// --- Siemens Structured Format ---
DATA_BLOCK "model__HS16_IW50_"
{ S7_Optimized_Access := 'TRUE' }
VERSION :
NON_RETAIN
   VAR
      W_i : ARRAY[0..15, 0..39] OF REAL;
      W_f : ARRAY[0..15, 0..39] OF REAL;
      W_g : ARRAY[0..15, 0..39] OF REAL;
      W_o : ARRAY[0..15, 0..39] OF REAL;
      R_i : ARRAY[0..15, 0..15] OF REAL;
      R_f : ARRAY[0..15, 0..15] OF REAL;
      R_g : ARRAY[0..15, 0..15] OF REAL;
      R_o : ARRAY[0..15, 0..15] OF REAL;
      B_i : ARRAY[0..15] OF REAL;
      B_f : ARRAY[0..15] OF REAL;
      B_g : ARRAY[0..15] OF REAL;
      B_o : ARRAY[0..15] OF REAL;
      FC_W : ARRAY[0..39, 0..15] OF REAL;
      FC_B : ARRAY[0..39] OF REAL;
   END_VAR
BEGIN

      W_i[0,0] := -0.02612339;
      W_i[0,1] := 0.12072767;
      W_i[0,2] := -0.02244412;
      W_i[0,3] := -0.02933176;
      W_i[0,4] := 0.13427743;
      W_i[0,5] := -0.01298498;
      W_i[0,6] := -0.08133418;
      W_i[0,7] := 0.19622199;
      W_i[0,8] := 0.14236863;
      W_i[0,9] := -0.06801347;
      W_i[0,10] := 0.16722029;
      W_i[0,11] := -0.33964941;
      W_i[0,12] := -0.82021421;
      W_i[0,13] := 0.06192777;
      W_i[0,14] := 0.39121246;
      W_i[0,15] := -0.96388686;
      W_i[0,16] := 0.14144035;
      W_i[0,17] := -0.25961453;
      W_i[0,18] := 0.00280210;
      W_i[0,19] := 0.36805412;
      W_i[0,20] := 0.11180947;
      W_i[0,21] := 0.28874406;
      W_i[0,22] := 0.24604218;
      W_i[0,23] := 0.06171668;
      W_i[0,24] := 0.88452333;
      W_i[0,25] := 0.96678102;
      W_i[0,26] := 0.04491860;
      W_i[0,27] := -0.21186443;
      W_i[0,28] := 0.08944755;
      W_i[0,29] := -0.10767028;
      W_i[0,30] := 0.60365808;
      W_i[0,31] := -0.13146588;
      W_i[0,32] := 0.12239406;
      W_i[0,33] := -0.09614152;
      W_i[0,34] := 1.05674243;
      W_i[0,35] := -0.04317053;
      W_i[0,36] := 0.15985158;
      W_i[0,37] := -0.00158236;
      W_i[0,38] := 0.64556688;
      W_i[0,39] := 0.15716811;
      W_i[1,0] := 0.02739522;
      W_i[1,1] := 0.10316847;
      W_i[1,2] := 0.01493799;
      W_i[1,3] := 0.01172978;
      W_i[1,4] := 0.17755681;
      W_i[1,5] := 0.02642176;
      W_i[1,6] := 0.08478273;
      W_i[1,7] := 0.04226714;
      W_i[1,8] := 0.00695325;
      W_i[1,9] := 0.03251113;
      W_i[1,10] := 0.02126005;
      W_i[1,11] := -0.01568736;
      W_i[1,12] := -0.09019557;
      W_i[1,13] := -0.08720633;
      W_i[1,14] := 0.02817911;
      W_i[1,15] := -0.01798955;
      W_i[1,16] := -0.04418186;
      W_i[1,17] := 0.01428624;
      W_i[1,18] := -0.27951232;
      W_i[1,19] := 0.05315392;
      W_i[1,20] := -0.10911061;
      W_i[1,21] := 0.05054765;
      W_i[1,22] := 0.18948558;
      W_i[1,23] := -0.08133697;
      W_i[1,24] := -0.40616348;
      W_i[1,25] := -0.53565234;
      W_i[1,26] := -0.10580445;
      W_i[1,27] := -0.17574981;
      W_i[1,28] := -0.05870668;
      W_i[1,29] := 0.05139971;
      W_i[1,30] := 0.03107365;
      W_i[1,31] := -0.09318750;
      W_i[1,32] := -0.25166753;
      W_i[1,33] := -0.11112119;
      W_i[1,34] := 0.15034710;
      W_i[1,35] := -0.26474807;
      W_i[1,36] := -0.05716439;
      W_i[1,37] := -0.00181797;
      W_i[1,38] := 0.06692428;
      W_i[1,39] := -0.00409455;
      W_i[2,0] := -0.04371461;
      W_i[2,1] := 0.03530892;
      W_i[2,2] := -0.03434504;
      W_i[2,3] := -0.05561700;
      W_i[2,4] := 0.00493065;
      W_i[2,5] := 0.03415375;
      W_i[2,6] := -0.02065521;
      W_i[2,7] := -0.04744798;
      W_i[2,8] := 0.11951899;
      W_i[2,9] := 0.11182401;
      W_i[2,10] := 0.04235537;
      W_i[2,11] := -0.08501492;
      W_i[2,12] := 0.08836282;
      W_i[2,13] := -0.03698122;
      W_i[2,14] := 0.11667735;
      W_i[2,15] := -1.35210800;
      W_i[2,16] := 0.04032730;
      W_i[2,17] := 0.39463934;
      W_i[2,18] := 0.23274027;
      W_i[2,19] := -0.09035096;
      W_i[2,20] := 0.02598169;
      W_i[2,21] := -0.02158709;
      W_i[2,22] := 0.08459560;
      W_i[2,23] := -0.01336102;
      W_i[2,24] := 0.39533728;
      W_i[2,25] := 0.21617500;
      W_i[2,26] := 0.04206325;
      W_i[2,27] := 0.03110088;
      W_i[2,28] := 0.00954145;
      W_i[2,29] := -0.08245377;
      W_i[2,30] := -0.01272953;
      W_i[2,31] := -0.00777793;
      W_i[2,32] := -0.03093930;
      W_i[2,33] := -0.14403637;
      W_i[2,34] := -0.36296284;
      W_i[2,35] := 0.02933266;
      W_i[2,36] := 0.00311332;
      W_i[2,37] := 0.06835733;
      W_i[2,38] := 0.13729195;
      W_i[2,39] := -0.09952185;
      W_i[3,0] := 0.00846558;
      W_i[3,1] := -0.12918584;
      W_i[3,2] := -0.00730979;
      W_i[3,3] := 0.01713126;
      W_i[3,4] := -0.02458502;
      W_i[3,5] := -0.01639076;
      W_i[3,6] := -0.17934421;
      W_i[3,7] := -0.01638387;
      W_i[3,8] := -0.03064539;
      W_i[3,9] := 0.08878898;
      W_i[3,10] := -0.07486653;
      W_i[3,11] := -0.08080578;
      W_i[3,12] := 0.06557790;
      W_i[3,13] := 0.01592479;
      W_i[3,14] := -0.03430796;
      W_i[3,15] := 0.01604570;
      W_i[3,16] := 0.01997751;
      W_i[3,17] := -0.03321569;
      W_i[3,18] := 0.04693119;
      W_i[3,19] := 0.00119276;
      W_i[3,20] := -0.06343115;
      W_i[3,21] := 0.07300727;
      W_i[3,22] := 0.17427416;
      W_i[3,23] := -0.07701004;
      W_i[3,24] := -0.04349097;
      W_i[3,25] := 0.08956601;
      W_i[3,26] := -0.03523625;
      W_i[3,27] := -0.00686803;
      W_i[3,28] := -0.01029908;
      W_i[3,29] := 0.05175918;
      W_i[3,30] := 0.10149232;
      W_i[3,31] := -0.11382963;
      W_i[3,32] := 0.07062076;
      W_i[3,33] := -0.01815722;
      W_i[3,34] := 0.04715188;
      W_i[3,35] := -0.06669057;
      W_i[3,36] := 0.01020681;
      W_i[3,37] := 0.25148758;
      W_i[3,38] := -0.01007098;
      W_i[3,39] := -0.00052197;
      W_i[4,0] := 0.06882605;
      W_i[4,1] := 0.29223976;
      W_i[4,2] := 0.13380581;
      W_i[4,3] := -0.35771182;
      W_i[4,4] := 0.25656733;
      W_i[4,5] := -0.20841958;
      W_i[4,6] := 0.07243224;
      W_i[4,7] := 0.38866916;
      W_i[4,8] := 0.53406250;
      W_i[4,9] := -0.23149215;
      W_i[4,10] := -0.19491005;
      W_i[4,11] := -0.48210201;
      W_i[4,12] := 0.13137554;
      W_i[4,13] := 0.50133437;
      W_i[4,14] := -0.01319221;
      W_i[4,15] := -0.16763180;
      W_i[4,16] := -0.02528067;
      W_i[4,17] := 0.20047617;
      W_i[4,18] := 0.07556880;
      W_i[4,19] := 0.12009662;
      W_i[4,20] := -0.23959216;
      W_i[4,21] := -0.05043668;
      W_i[4,22] := 0.03819416;
      W_i[4,23] := 0.32712597;
      W_i[4,24] := -0.06839418;
      W_i[4,25] := -0.00276239;
      W_i[4,26] := -0.26127121;
      W_i[4,27] := -0.20213830;
      W_i[4,28] := 0.07294428;
      W_i[4,29] := 0.04953664;
      W_i[4,30] := -0.04174086;
      W_i[4,31] := -0.06637315;
      W_i[4,32] := 0.09226974;
      W_i[4,33] := 0.13355142;
      W_i[4,34] := 0.09484247;
      W_i[4,35] := -0.09734286;
      W_i[4,36] := 0.03169553;
      W_i[4,37] := -0.08991057;
      W_i[4,38] := -0.13476068;
      W_i[4,39] := 0.29272395;
      W_i[5,0] := -0.05475799;
      W_i[5,1] := -0.06864791;
      W_i[5,2] := -0.02113621;
      W_i[5,3] := 0.02720109;
      W_i[5,4] := 0.10207788;
      W_i[5,5] := -0.00895342;
      W_i[5,6] := -0.02244009;
      W_i[5,7] := 0.16509427;
      W_i[5,8] := 0.01703463;
      W_i[5,9] := -0.21540523;
      W_i[5,10] := -0.00765499;
      W_i[5,11] := 0.01468746;
      W_i[5,12] := 0.22010665;
      W_i[5,13] := -0.09001971;
      W_i[5,14] := -0.02117113;
      W_i[5,15] := 0.07194266;
      W_i[5,16] := -0.18253084;
      W_i[5,17] := 0.04095849;
      W_i[5,18] := -0.08197289;
      W_i[5,19] := -0.27980739;
      W_i[5,20] := 0.11807738;
      W_i[5,21] := 0.25605229;
      W_i[5,22] := -0.18898037;
      W_i[5,23] := 0.06701536;
      W_i[5,24] := -0.38402686;
      W_i[5,25] := 0.03199298;
      W_i[5,26] := 0.28137541;
      W_i[5,27] := -0.03393725;
      W_i[5,28] := -0.00611741;
      W_i[5,29] := -0.21439074;
      W_i[5,30] := -0.24789658;
      W_i[5,31] := 0.01456884;
      W_i[5,32] := 0.09658974;
      W_i[5,33] := 0.07787250;
      W_i[5,34] := -0.00873361;
      W_i[5,35] := 0.02078887;
      W_i[5,36] := -0.00982943;
      W_i[5,37] := -0.22429584;
      W_i[5,38] := 0.25736400;
      W_i[5,39] := -0.30378288;
      W_i[6,0] := -0.15429787;
      W_i[6,1] := -0.00725780;
      W_i[6,2] := -0.01294193;
      W_i[6,3] := -0.08215277;
      W_i[6,4] := -0.13259856;
      W_i[6,5] := -0.16592383;
      W_i[6,6] := -0.00615384;
      W_i[6,7] := 0.02707914;
      W_i[6,8] := 0.03321055;
      W_i[6,9] := 0.20581089;
      W_i[6,10] := -0.02888039;
      W_i[6,11] := 0.13899046;
      W_i[6,12] := -0.50004631;
      W_i[6,13] := -0.18613359;
      W_i[6,14] := 0.02271620;
      W_i[6,15] := -0.05991226;
      W_i[6,16] := 0.02941754;
      W_i[6,17] := -0.05727729;
      W_i[6,18] := -0.05220168;
      W_i[6,19] := 0.12824084;
      W_i[6,20] := -0.11432266;
      W_i[6,21] := -0.06927077;
      W_i[6,22] := -0.16510975;
      W_i[6,23] := 0.16503085;
      W_i[6,24] := -0.06193599;
      W_i[6,25] := 0.08007926;
      W_i[6,26] := 0.16539313;
      W_i[6,27] := -0.09439778;
      W_i[6,28] := -0.11654797;
      W_i[6,29] := -0.07672822;
      W_i[6,30] := -0.09051897;
      W_i[6,31] := -0.05891651;
      W_i[6,32] := -0.06850113;
      W_i[6,33] := -0.01238405;
      W_i[6,34] := 0.05435950;
      W_i[6,35] := -0.07693552;
      W_i[6,36] := 0.00911314;
      W_i[6,37] := -0.01921199;
      W_i[6,38] := 0.05525052;
      W_i[6,39] := -0.07226433;
      W_i[7,0] := -0.19423574;
      W_i[7,1] := -0.24973391;
      W_i[7,2] := -0.05149378;
      W_i[7,3] := -0.25323981;
      W_i[7,4] := 0.39798826;
      W_i[7,5] := 0.24827355;
      W_i[7,6] := 0.43568289;
      W_i[7,7] := -0.13336283;
      W_i[7,8] := 0.12423158;
      W_i[7,9] := -0.07743893;
      W_i[7,10] := -0.15183467;
      W_i[7,11] := 0.06914197;
      W_i[7,12] := -0.02671312;
      W_i[7,13] := -0.21586929;
      W_i[7,14] := 0.00868284;
      W_i[7,15] := 0.02255189;
      W_i[7,16] := -0.02795821;
      W_i[7,17] := 0.00887333;
      W_i[7,18] := -0.12309828;
      W_i[7,19] := -0.00309656;
      W_i[7,20] := 0.38424814;
      W_i[7,21] := 0.30607188;
      W_i[7,22] := -0.15942656;
      W_i[7,23] := 0.01897525;
      W_i[7,24] := -0.09797664;
      W_i[7,25] := -0.02867761;
      W_i[7,26] := 0.15050705;
      W_i[7,27] := 0.00785798;
      W_i[7,28] := -0.19198960;
      W_i[7,29] := 0.21648924;
      W_i[7,30] := 0.16888635;
      W_i[7,31] := -0.00119574;
      W_i[7,32] := -0.24025443;
      W_i[7,33] := 0.30170068;
      W_i[7,34] := 0.23723993;
      W_i[7,35] := -0.13449760;
      W_i[7,36] := -0.15990667;
      W_i[7,37] := -0.00520837;
      W_i[7,38] := 0.08311661;
      W_i[7,39] := -0.02735133;
      W_i[8,0] := -0.06984207;
      W_i[8,1] := 0.18467268;
      W_i[8,2] := 0.00678134;
      W_i[8,3] := 0.04922282;
      W_i[8,4] := 0.11598286;
      W_i[8,5] := 0.08822776;
      W_i[8,6] := -0.10902181;
      W_i[8,7] := -0.16074504;
      W_i[8,8] := -0.11118431;
      W_i[8,9] := 0.10051250;
      W_i[8,10] := 0.07012353;
      W_i[8,11] := 0.07681172;
      W_i[8,12] := -0.22344230;
      W_i[8,13] := -0.12049098;
      W_i[8,14] := 0.01157948;
      W_i[8,15] := 0.01269015;
      W_i[8,16] := 0.01600377;
      W_i[8,17] := 0.02240872;
      W_i[8,18] := -0.02060430;
      W_i[8,19] := -0.06097650;
      W_i[8,20] := 0.07957297;
      W_i[8,21] := 0.08196621;
      W_i[8,22] := -0.02732777;
      W_i[8,23] := -0.06837825;
      W_i[8,24] := -1.24913669;
      W_i[8,25] := -0.21292350;
      W_i[8,26] := 0.05969907;
      W_i[8,27] := -0.15808001;
      W_i[8,28] := -0.06865929;
      W_i[8,29] := -0.05003216;
      W_i[8,30] := 0.13252324;
      W_i[8,31] := -0.10141694;
      W_i[8,32] := 0.15883078;
      W_i[8,33] := 0.01671924;
      W_i[8,34] := 0.01595451;
      W_i[8,35] := 0.04233614;
      W_i[8,36] := 0.10780733;
      W_i[8,37] := 0.00896461;
      W_i[8,38] := 0.13257688;
      W_i[8,39] := 0.05639813;
      W_i[9,0] := 0.04840493;
      W_i[9,1] := 0.00527499;
      W_i[9,2] := -0.03278387;
      W_i[9,3] := 0.08216210;
      W_i[9,4] := -0.01587271;
      W_i[9,5] := -0.00737574;
      W_i[9,6] := -0.01856831;
      W_i[9,7] := 0.19069298;
      W_i[9,8] := -0.00912018;
      W_i[9,9] := -0.24746008;
      W_i[9,10] := -0.06627475;
      W_i[9,11] := 0.07460143;
      W_i[9,12] := -0.04468247;
      W_i[9,13] := -0.03485956;
      W_i[9,14] := -0.02453788;
      W_i[9,15] := 0.00244658;
      W_i[9,16] := -0.00826298;
      W_i[9,17] := 0.00922262;
      W_i[9,18] := 0.03385285;
      W_i[9,19] := 0.04683683;
      W_i[9,20] := -0.03658741;
      W_i[9,21] := -0.05278853;
      W_i[9,22] := -0.06786657;
      W_i[9,23] := -0.03328852;
      W_i[9,24] := -0.67544466;
      W_i[9,25] := -0.45174205;
      W_i[9,26] := 0.01428142;
      W_i[9,27] := 0.00258533;
      W_i[9,28] := -0.00212107;
      W_i[9,29] := 0.26447642;
      W_i[9,30] := -0.04738332;
      W_i[9,31] := 0.02417716;
      W_i[9,32] := -0.13879688;
      W_i[9,33] := 0.05013292;
      W_i[9,34] := -0.61316240;
      W_i[9,35] := -0.11345586;
      W_i[9,36] := -0.00836167;
      W_i[9,37] := 0.06233503;
      W_i[9,38] := -0.01308454;
      W_i[9,39] := 0.00902628;
      W_i[10,0] := 0.05447512;
      W_i[10,1] := 0.00135808;
      W_i[10,2] := 0.00598898;
      W_i[10,3] := -0.00021247;
      W_i[10,4] := 0.00281035;
      W_i[10,5] := -0.01504579;
      W_i[10,6] := 0.12122837;
      W_i[10,7] := -0.06385819;
      W_i[10,8] := -0.04342161;
      W_i[10,9] := 0.08000173;
      W_i[10,10] := 0.01194646;
      W_i[10,11] := 0.11263964;
      W_i[10,12] := 0.04725603;
      W_i[10,13] := -0.02525371;
      W_i[10,14] := 0.01381323;
      W_i[10,15] := 0.00554248;
      W_i[10,16] := -0.01660426;
      W_i[10,17] := 0.00241101;
      W_i[10,18] := 0.01211567;
      W_i[10,19] := 0.01751081;
      W_i[10,20] := -0.00082530;
      W_i[10,21] := 0.03101674;
      W_i[10,22] := -0.26447886;
      W_i[10,23] := 0.02353600;
      W_i[10,24] := -0.22910219;
      W_i[10,25] := -0.38894618;
      W_i[10,26] := -0.03487613;
      W_i[10,27] := -0.11107682;
      W_i[10,28] := -0.06958691;
      W_i[10,29] := 0.15007824;
      W_i[10,30] := 0.10014386;
      W_i[10,31] := 0.07397891;
      W_i[10,32] := -0.12383275;
      W_i[10,33] := 0.08686586;
      W_i[10,34] := -0.85524035;
      W_i[10,35] := 0.14177939;
      W_i[10,36] := -0.02201772;
      W_i[10,37] := 0.01626217;
      W_i[10,38] := 0.16784185;
      W_i[10,39] := 0.00716509;
      W_i[11,0] := -0.08976970;
      W_i[11,1] := -0.00744615;
      W_i[11,2] := -0.05819619;
      W_i[11,3] := -0.07143553;
      W_i[11,4] := -0.03154673;
      W_i[11,5] := 0.03580843;
      W_i[11,6] := -0.03945105;
      W_i[11,7] := -0.12150279;
      W_i[11,8] := 0.00981623;
      W_i[11,9] := 0.05031164;
      W_i[11,10] := -0.02300070;
      W_i[11,11] := -0.08073328;
      W_i[11,12] := 0.01272614;
      W_i[11,13] := -0.07925726;
      W_i[11,14] := 0.00678512;
      W_i[11,15] := 0.04620445;
      W_i[11,16] := -0.00129330;
      W_i[11,17] := 0.00041449;
      W_i[11,18] := 0.03960210;
      W_i[11,19] := -0.01602606;
      W_i[11,20] := 0.02149412;
      W_i[11,21] := -0.02751144;
      W_i[11,22] := -0.15877301;
      W_i[11,23] := 0.01397473;
      W_i[11,24] := -0.66238141;
      W_i[11,25] := -0.94520783;
      W_i[11,26] := -0.10410358;
      W_i[11,27] := -0.01858253;
      W_i[11,28] := -0.07172703;
      W_i[11,29] := 0.25134814;
      W_i[11,30] := -0.14801161;
      W_i[11,31] := -0.01742411;
      W_i[11,32] := 0.07450388;
      W_i[11,33] := -0.03559265;
      W_i[11,34] := -0.21006276;
      W_i[11,35] := 0.20278554;
      W_i[11,36] := -0.01763817;
      W_i[11,37] := -0.27180666;
      W_i[11,38] := 0.05380114;
      W_i[11,39] := 0.00796253;
      W_i[12,0] := 0.25864720;
      W_i[12,1] := -0.12210964;
      W_i[12,2] := -0.14704542;
      W_i[12,3] := -0.03986358;
      W_i[12,4] := 0.08733799;
      W_i[12,5] := -0.37284544;
      W_i[12,6] := 0.10571802;
      W_i[12,7] := -0.11933661;
      W_i[12,8] := -0.06846283;
      W_i[12,9] := 0.08954131;
      W_i[12,10] := -0.22306511;
      W_i[12,11] := 0.46803057;
      W_i[12,12] := 0.21598789;
      W_i[12,13] := -0.09787964;
      W_i[12,14] := 0.15112200;
      W_i[12,15] := 0.20643055;
      W_i[12,16] := -0.07569909;
      W_i[12,17] := -0.00754971;
      W_i[12,18] := -0.09548484;
      W_i[12,19] := 0.01058478;
      W_i[12,20] := 0.47774643;
      W_i[12,21] := -0.12664053;
      W_i[12,22] := 0.20265566;
      W_i[12,23] := 0.19177310;
      W_i[12,24] := 0.31017169;
      W_i[12,25] := 0.23971170;
      W_i[12,26] := -0.31540856;
      W_i[12,27] := 0.03726046;
      W_i[12,28] := -0.08490968;
      W_i[12,29] := 0.18619052;
      W_i[12,30] := 0.18660802;
      W_i[12,31] := -0.07303433;
      W_i[12,32] := 0.10245761;
      W_i[12,33] := -0.12202786;
      W_i[12,34] := -0.00883020;
      W_i[12,35] := -0.27889481;
      W_i[12,36] := 0.19747989;
      W_i[12,37] := -0.33369049;
      W_i[12,38] := 0.28634214;
      W_i[12,39] := 0.08568040;
      W_i[13,0] := -0.12176741;
      W_i[13,1] := 0.13172998;
      W_i[13,2] := -0.01483796;
      W_i[13,3] := -0.02370377;
      W_i[13,4] := 0.14033392;
      W_i[13,5] := -0.02840229;
      W_i[13,6] := -0.06477696;
      W_i[13,7] := -0.09099311;
      W_i[13,8] := -0.02282218;
      W_i[13,9] := 0.24101490;
      W_i[13,10] := 0.02915199;
      W_i[13,11] := -0.20095268;
      W_i[13,12] := -0.41396245;
      W_i[13,13] := -0.09245090;
      W_i[13,14] := 0.02569151;
      W_i[13,15] := -0.04253404;
      W_i[13,16] := -0.03762357;
      W_i[13,17] := 0.03585879;
      W_i[13,18] := 0.01942859;
      W_i[13,19] := 0.13924608;
      W_i[13,20] := 0.02253839;
      W_i[13,21] := 0.04408298;
      W_i[13,22] := 0.11049129;
      W_i[13,23] := 0.09530613;
      W_i[13,24] := 0.22805369;
      W_i[13,25] := -0.03002743;
      W_i[13,26] := 0.14904597;
      W_i[13,27] := 0.04909040;
      W_i[13,28] := -0.01216692;
      W_i[13,29] := -0.08759474;
      W_i[13,30] := 0.09012819;
      W_i[13,31] := -0.05122391;
      W_i[13,32] := -0.07538325;
      W_i[13,33] := 0.01453052;
      W_i[13,34] := -0.06318332;
      W_i[13,35] := -0.08720891;
      W_i[13,36] := 0.07678616;
      W_i[13,37] := 0.13920598;
      W_i[13,38] := -0.06368222;
      W_i[13,39] := 1.11653936;
      W_i[14,0] := -0.07855019;
      W_i[14,1] := 0.03459382;
      W_i[14,2] := -0.02766559;
      W_i[14,3] := 0.04799297;
      W_i[14,4] := 0.02599700;
      W_i[14,5] := 0.06535108;
      W_i[14,6] := 0.00835573;
      W_i[14,7] := -0.06900378;
      W_i[14,8] := -0.02075530;
      W_i[14,9] := 0.05139967;
      W_i[14,10] := 0.01833898;
      W_i[14,11] := -0.09905620;
      W_i[14,12] := 0.04986498;
      W_i[14,13] := 0.08562920;
      W_i[14,14] := 0.04875882;
      W_i[14,15] := 0.21624923;
      W_i[14,16] := -0.09095794;
      W_i[14,17] := -0.00323463;
      W_i[14,18] := 0.52891386;
      W_i[14,19] := -0.31447127;
      W_i[14,20] := 0.04405079;
      W_i[14,21] := -0.04545887;
      W_i[14,22] := -0.18876931;
      W_i[14,23] := -0.04623262;
      W_i[14,24] := -0.37235597;
      W_i[14,25] := -0.34788635;
      W_i[14,26] := -0.16801551;
      W_i[14,27] := 0.07317468;
      W_i[14,28] := 0.02443709;
      W_i[14,29] := 0.24874535;
      W_i[14,30] := -0.39551601;
      W_i[14,31] := -0.07593500;
      W_i[14,32] := -0.28626809;
      W_i[14,33] := -0.31125993;
      W_i[14,34] := -0.64042038;
      W_i[14,35] := 0.03362265;
      W_i[14,36] := 0.02987647;
      W_i[14,37] := -0.11912733;
      W_i[14,38] := 0.20975146;
      W_i[14,39] := 0.74268162;
      W_i[15,0] := 0.05764041;
      W_i[15,1] := 0.01238812;
      W_i[15,2] := -0.00211884;
      W_i[15,3] := -0.15071799;
      W_i[15,4] := -0.05083022;
      W_i[15,5] := 0.03901526;
      W_i[15,6] := -0.02054744;
      W_i[15,7] := 0.00484566;
      W_i[15,8] := 0.03377596;
      W_i[15,9] := 0.06261286;
      W_i[15,10] := 0.02025893;
      W_i[15,11] := 0.09115529;
      W_i[15,12] := 0.02875202;
      W_i[15,13] := 0.02998743;
      W_i[15,14] := -0.00594068;
      W_i[15,15] := -0.01918536;
      W_i[15,16] := -0.01136775;
      W_i[15,17] := 0.00490831;
      W_i[15,18] := -0.07127053;
      W_i[15,19] := -0.02636776;
      W_i[15,20] := 0.06915537;
      W_i[15,21] := 0.25859579;
      W_i[15,22] := -0.39175701;
      W_i[15,23] := 0.03068081;
      W_i[15,24] := -0.66952252;
      W_i[15,25] := -0.82186484;
      W_i[15,26] := 0.00559764;
      W_i[15,27] := -0.04806713;
      W_i[15,28] := -0.05927165;
      W_i[15,29] := -0.02447721;
      W_i[15,30] := -0.35062087;
      W_i[15,31] := -0.01519912;
      W_i[15,32] := -0.12022296;
      W_i[15,33] := 0.17821504;
      W_i[15,34] := -0.81185091;
      W_i[15,35] := -0.22858475;
      W_i[15,36] := -0.06415448;
      W_i[15,37] := -0.17577237;
      W_i[15,38] := 0.00998123;
      W_i[15,39] := 0.04287737;
      W_f[0,0] := 0.04715263;
      W_f[0,1] := 0.10899676;
      W_f[0,2] := -0.06567381;
      W_f[0,3] := 0.08125947;
      W_f[0,4] := -0.12792981;
      W_f[0,5] := 0.02464872;
      W_f[0,6] := -0.00594598;
      W_f[0,7] := 0.00857108;
      W_f[0,8] := -0.02990395;
      W_f[0,9] := -0.03421510;
      W_f[0,10] := 0.10801075;
      W_f[0,11] := -0.16118450;
      W_f[0,12] := 0.06628553;
      W_f[0,13] := -0.00627413;
      W_f[0,14] := -0.09413274;
      W_f[0,15] := -0.02655103;
      W_f[0,16] := 0.04184651;
      W_f[0,17] := -0.13916989;
      W_f[0,18] := -0.11053458;
      W_f[0,19] := -0.15861273;
      W_f[0,20] := 0.03201112;
      W_f[0,21] := 0.19275719;
      W_f[0,22] := 0.27139077;
      W_f[0,23] := -0.01148643;
      W_f[0,24] := 0.96007264;
      W_f[0,25] := 0.87839752;
      W_f[0,26] := -0.03665132;
      W_f[0,27] := -0.01417279;
      W_f[0,28] := -0.03944051;
      W_f[0,29] := -0.21950646;
      W_f[0,30] := 0.28375676;
      W_f[0,31] := 0.06307220;
      W_f[0,32] := 0.33201745;
      W_f[0,33] := 0.12054460;
      W_f[0,34] := 0.68658948;
      W_f[0,35] := 0.23550873;
      W_f[0,36] := -0.01086835;
      W_f[0,37] := -0.08451042;
      W_f[0,38] := -0.00964221;
      W_f[0,39] := -0.03436853;
      W_f[1,0] := 0.08623593;
      W_f[1,1] := -0.73259664;
      W_f[1,2] := 0.08433209;
      W_f[1,3] := -0.03844298;
      W_f[1,4] := -0.11556439;
      W_f[1,5] := 0.20516349;
      W_f[1,6] := -0.10453314;
      W_f[1,7] := -0.04163654;
      W_f[1,8] := -0.04797882;
      W_f[1,9] := -0.06256276;
      W_f[1,10] := -0.09822980;
      W_f[1,11] := 0.12738556;
      W_f[1,12] := 0.23426814;
      W_f[1,13] := 0.09855855;
      W_f[1,14] := 0.03435090;
      W_f[1,15] := 0.11293387;
      W_f[1,16] := -0.19483942;
      W_f[1,17] := -0.03186984;
      W_f[1,18] := 0.66178006;
      W_f[1,19] := 0.02745492;
      W_f[1,20] := 0.35740805;
      W_f[1,21] := -0.25831303;
      W_f[1,22] := -0.12126569;
      W_f[1,23] := 0.22377175;
      W_f[1,24] := -0.83024675;
      W_f[1,25] := -1.25248599;
      W_f[1,26] := 0.28189325;
      W_f[1,27] := -0.13919783;
      W_f[1,28] := -0.02240801;
      W_f[1,29] := -0.18801042;
      W_f[1,30] := -0.04805183;
      W_f[1,31] := 0.24313359;
      W_f[1,32] := 0.26400492;
      W_f[1,33] := 0.17501286;
      W_f[1,34] := 0.51169682;
      W_f[1,35] := 0.40932828;
      W_f[1,36] := -0.35491022;
      W_f[1,37] := -0.03798340;
      W_f[1,38] := -0.08608454;
      W_f[1,39] := 0.02175015;
      W_f[2,0] := -0.00661589;
      W_f[2,1] := -0.13814320;
      W_f[2,2] := 0.02391077;
      W_f[2,3] := 0.15640482;
      W_f[2,4] := 0.00755587;
      W_f[2,5] := -0.04414793;
      W_f[2,6] := -0.05434313;
      W_f[2,7] := 0.06549069;
      W_f[2,8] := -0.15011497;
      W_f[2,9] := -0.08841761;
      W_f[2,10] := 0.00392893;
      W_f[2,11] := 0.61885518;
      W_f[2,12] := 0.55919319;
      W_f[2,13] := 0.02260459;
      W_f[2,14] := -0.20439312;
      W_f[2,15] := 0.25819176;
      W_f[2,16] := 0.00852524;
      W_f[2,17] := 0.36273137;
      W_f[2,18] := -0.45172021;
      W_f[2,19] := 0.06631603;
      W_f[2,20] := 0.09949520;
      W_f[2,21] := 0.06160212;
      W_f[2,22] := -0.03724279;
      W_f[2,23] := -0.01405078;
      W_f[2,24] := -1.01044071;
      W_f[2,25] := -1.24477458;
      W_f[2,26] := 0.06317704;
      W_f[2,27] := -0.12849498;
      W_f[2,28] := -0.01733010;
      W_f[2,29] := 0.30296484;
      W_f[2,30] := -0.06890817;
      W_f[2,31] := 0.12288452;
      W_f[2,32] := 0.03147413;
      W_f[2,33] := 0.24991731;
      W_f[2,34] := 0.14598863;
      W_f[2,35] := -0.05373066;
      W_f[2,36] := -0.08683386;
      W_f[2,37] := 0.17713107;
      W_f[2,38] := -0.31477356;
      W_f[2,39] := 1.00106454;
      W_f[3,0] := -0.00357926;
      W_f[3,1] := -0.02668277;
      W_f[3,2] := -0.02272550;
      W_f[3,3] := 0.04566845;
      W_f[3,4] := -0.05781303;
      W_f[3,5] := -0.05116368;
      W_f[3,6] := 0.33208069;
      W_f[3,7] := 0.05969469;
      W_f[3,8] := 0.04631799;
      W_f[3,9] := -0.07284315;
      W_f[3,10] := 0.02255991;
      W_f[3,11] := 0.05159385;
      W_f[3,12] := -0.20268613;
      W_f[3,13] := 0.01119571;
      W_f[3,14] := -0.05706387;
      W_f[3,15] := -0.07039116;
      W_f[3,16] := 0.01233673;
      W_f[3,17] := -0.11033136;
      W_f[3,18] := 0.03755057;
      W_f[3,19] := -0.15966073;
      W_f[3,20] := -0.00759900;
      W_f[3,21] := 0.02997555;
      W_f[3,22] := -0.00575700;
      W_f[3,23] := 0.09471051;
      W_f[3,24] := -0.76867020;
      W_f[3,25] := -1.10453773;
      W_f[3,26] := 0.08160409;
      W_f[3,27] := 0.07287289;
      W_f[3,28] := -0.23396601;
      W_f[3,29] := -0.01620052;
      W_f[3,30] := -0.14668229;
      W_f[3,31] := 0.29359242;
      W_f[3,32] := 0.28141207;
      W_f[3,33] := 0.10357075;
      W_f[3,34] := 0.15553899;
      W_f[3,35] := -0.08215727;
      W_f[3,36] := 0.59300834;
      W_f[3,37] := 0.06939243;
      W_f[3,38] := 0.05595111;
      W_f[3,39] := -0.01764361;
      W_f[4,0] := -0.04732760;
      W_f[4,1] := 0.14226569;
      W_f[4,2] := -0.19679488;
      W_f[4,3] := 0.03169706;
      W_f[4,4] := 0.03950732;
      W_f[4,5] := 0.12956409;
      W_f[4,6] := -0.13465910;
      W_f[4,7] := -0.11123411;
      W_f[4,8] := 0.01169378;
      W_f[4,9] := -0.00041270;
      W_f[4,10] := 0.06247496;
      W_f[4,11] := -0.19790170;
      W_f[4,12] := -0.13562107;
      W_f[4,13] := 0.40435797;
      W_f[4,14] := 0.03306964;
      W_f[4,15] := -0.17322055;
      W_f[4,16] := -0.05731088;
      W_f[4,17] := -0.06482833;
      W_f[4,18] := 0.09320654;
      W_f[4,19] := 0.24850778;
      W_f[4,20] := -0.18519133;
      W_f[4,21] := 0.12798916;
      W_f[4,22] := 0.14323689;
      W_f[4,23] := -0.01742595;
      W_f[4,24] := 1.63087487;
      W_f[4,25] := 1.71278691;
      W_f[4,26] := -0.17371880;
      W_f[4,27] := 0.04438495;
      W_f[4,28] := 0.10424647;
      W_f[4,29] := 0.17063302;
      W_f[4,30] := 0.42905927;
      W_f[4,31] := 0.27194634;
      W_f[4,32] := -0.01861881;
      W_f[4,33] := -0.02290395;
      W_f[4,34] := 0.25754037;
      W_f[4,35] := 0.41329530;
      W_f[4,36] := -0.09744941;
      W_f[4,37] := 0.27917421;
      W_f[4,38] := 0.01022570;
      W_f[4,39] := 0.21825342;
      W_f[5,0] := -0.12265578;
      W_f[5,1] := 0.11042612;
      W_f[5,2] := 0.03006834;
      W_f[5,3] := -0.26207334;
      W_f[5,4] := 0.00985776;
      W_f[5,5] := -0.02016665;
      W_f[5,6] := -0.03333576;
      W_f[5,7] := 0.15882950;
      W_f[5,8] := -0.27977559;
      W_f[5,9] := 0.25365406;
      W_f[5,10] := -0.03230783;
      W_f[5,11] := -0.21518956;
      W_f[5,12] := -0.23225260;
      W_f[5,13] := 0.04519130;
      W_f[5,14] := 0.00848376;
      W_f[5,15] := -0.03351771;
      W_f[5,16] := 0.09852035;
      W_f[5,17] := -0.09458777;
      W_f[5,18] := 0.02086790;
      W_f[5,19] := 0.13770969;
      W_f[5,20] := -0.04140184;
      W_f[5,21] := 0.09476180;
      W_f[5,22] := 0.41919291;
      W_f[5,23] := -0.14774488;
      W_f[5,24] := 1.13465798;
      W_f[5,25] := 1.46192527;
      W_f[5,26] := -0.06388761;
      W_f[5,27] := 0.03928265;
      W_f[5,28] := 0.03407076;
      W_f[5,29] := -0.51813745;
      W_f[5,30] := 0.24349271;
      W_f[5,31] := 0.01923511;
      W_f[5,32] := 0.05050964;
      W_f[5,33] := -0.03686145;
      W_f[5,34] := 1.16242385;
      W_f[5,35] := 0.04278161;
      W_f[5,36] := -0.03958681;
      W_f[5,37] := 0.17119792;
      W_f[5,38] := 0.04197992;
      W_f[5,39] := 0.22113459;
      W_f[6,0] := -0.05077897;
      W_f[6,1] := 0.12266269;
      W_f[6,2] := -0.15582716;
      W_f[6,3] := -0.07109610;
      W_f[6,4] := 0.01037609;
      W_f[6,5] := 0.03313427;
      W_f[6,6] := 0.05276644;
      W_f[6,7] := -0.06777491;
      W_f[6,8] := 0.02246877;
      W_f[6,9] := -0.12816820;
      W_f[6,10] := 0.01218652;
      W_f[6,11] := -0.06725728;
      W_f[6,12] := 0.11980707;
      W_f[6,13] := -0.03621849;
      W_f[6,14] := 0.23148635;
      W_f[6,15] := -0.05256491;
      W_f[6,16] := 0.28452423;
      W_f[6,17] := -0.04785041;
      W_f[6,18] := 0.00029584;
      W_f[6,19] := -0.33732000;
      W_f[6,20] := -0.01787652;
      W_f[6,21] := 0.04774499;
      W_f[6,22] := 0.32209477;
      W_f[6,23] := -0.11889420;
      W_f[6,24] := 1.09117067;
      W_f[6,25] := 1.12744486;
      W_f[6,26] := -0.07003234;
      W_f[6,27] := 0.01855475;
      W_f[6,28] := -0.00330310;
      W_f[6,29] := -0.26430756;
      W_f[6,30] := 0.21318698;
      W_f[6,31] := 0.04353658;
      W_f[6,32] := 0.27845708;
      W_f[6,33] := 0.02148022;
      W_f[6,34] := 1.27716565;
      W_f[6,35] := -0.13685782;
      W_f[6,36] := -0.05482837;
      W_f[6,37] := 0.09329895;
      W_f[6,38] := 0.06903394;
      W_f[6,39] := -0.18291597;
      W_f[7,0] := -0.06782078;
      W_f[7,1] := -0.41273677;
      W_f[7,2] := -0.23223357;
      W_f[7,3] := -0.13132100;
      W_f[7,4] := -0.00691312;
      W_f[7,5] := 0.61953580;
      W_f[7,6] := 0.74713135;
      W_f[7,7] := -0.13415965;
      W_f[7,8] := -0.70239842;
      W_f[7,9] := -0.12314104;
      W_f[7,10] := -0.26408386;
      W_f[7,11] := -0.04327460;
      W_f[7,12] := 0.06000946;
      W_f[7,13] := -0.08953854;
      W_f[7,14] := -0.01992717;
      W_f[7,15] := -0.03414788;
      W_f[7,16] := -0.10218910;
      W_f[7,17] := -0.02195402;
      W_f[7,18] := -0.15076502;
      W_f[7,19] := -0.14730737;
      W_f[7,20] := 0.04946668;
      W_f[7,21] := 0.36726916;
      W_f[7,22] := -0.01913268;
      W_f[7,23] := -0.20478757;
      W_f[7,24] := -0.07383893;
      W_f[7,25] := 0.03577507;
      W_f[7,26] := -0.36156556;
      W_f[7,27] := 0.10162932;
      W_f[7,28] := 0.08031812;
      W_f[7,29] := 0.03659641;
      W_f[7,30] := -0.06054391;
      W_f[7,31] := 0.01948766;
      W_f[7,32] := 0.22690910;
      W_f[7,33] := 0.09243126;
      W_f[7,34] := 0.36665705;
      W_f[7,35] := -0.18836242;
      W_f[7,36] := 0.08979291;
      W_f[7,37] := -0.03466015;
      W_f[7,38] := 0.17328687;
      W_f[7,39] := 0.01111504;
      W_f[8,0] := -0.10757597;
      W_f[8,1] := 0.18080002;
      W_f[8,2] := -0.18117517;
      W_f[8,3] := 0.05444926;
      W_f[8,4] := -0.03406826;
      W_f[8,5] := 0.03211219;
      W_f[8,6] := 0.04893153;
      W_f[8,7] := 0.00879812;
      W_f[8,8] := 0.05938864;
      W_f[8,9] := -0.05662099;
      W_f[8,10] := 0.05257615;
      W_f[8,11] := -0.27383971;
      W_f[8,12] := -0.06582582;
      W_f[8,13] := 0.00902832;
      W_f[8,14] := 0.01648709;
      W_f[8,15] := -0.32319725;
      W_f[8,16] := 0.18786642;
      W_f[8,17] := -0.08832575;
      W_f[8,18] := 0.05050201;
      W_f[8,19] := -0.14431089;
      W_f[8,20] := -0.07567763;
      W_f[8,21] := -0.01289035;
      W_f[8,22] := -0.01249675;
      W_f[8,23] := -0.01680613;
      W_f[8,24] := 0.68140340;
      W_f[8,25] := 0.89507484;
      W_f[8,26] := -0.06418619;
      W_f[8,27] := 0.07647979;
      W_f[8,28] := 0.03661409;
      W_f[8,29] := -0.14417614;
      W_f[8,30] := -0.04263573;
      W_f[8,31] := 0.03779473;
      W_f[8,32] := 0.05052606;
      W_f[8,33] := 0.06155790;
      W_f[8,34] := 1.02400410;
      W_f[8,35] := -0.17263915;
      W_f[8,36] := 0.00310001;
      W_f[8,37] := -0.04516594;
      W_f[8,38] := -0.01715083;
      W_f[8,39] := 0.20146139;
      W_f[9,0] := 0.15622687;
      W_f[9,1] := 0.10635939;
      W_f[9,2] := -0.72994000;
      W_f[9,3] := -0.14118610;
      W_f[9,4] := -0.14285882;
      W_f[9,5] := 0.16976678;
      W_f[9,6] := 0.04101548;
      W_f[9,7] := 0.27330139;
      W_f[9,8] := -0.28499794;
      W_f[9,9] := -0.18460013;
      W_f[9,10] := 0.00495566;
      W_f[9,11] := -0.10320173;
      W_f[9,12] := -0.06923575;
      W_f[9,13] := 0.01051456;
      W_f[9,14] := -0.04837225;
      W_f[9,15] := -0.07643475;
      W_f[9,16] := 0.09923542;
      W_f[9,17] := -0.00375771;
      W_f[9,18] := -0.02745963;
      W_f[9,19] := 0.00053912;
      W_f[9,20] := -0.08774224;
      W_f[9,21] := 0.14884678;
      W_f[9,22] := 0.02246397;
      W_f[9,23] := 0.02559338;
      W_f[9,24] := -0.25594050;
      W_f[9,25] := -0.34410420;
      W_f[9,26] := 0.00826990;
      W_f[9,27] := -0.00619870;
      W_f[9,28] := 0.02722283;
      W_f[9,29] := -0.04649381;
      W_f[9,30] := 0.32932112;
      W_f[9,31] := -0.01646173;
      W_f[9,32] := 0.16043368;
      W_f[9,33] := 0.15029813;
      W_f[9,34] := -0.59800792;
      W_f[9,35] := 0.31481645;
      W_f[9,36] := -0.03954235;
      W_f[9,37] := -0.10088660;
      W_f[9,38] := 0.07048618;
      W_f[9,39] := -0.02868455;
      W_f[10,0] := -0.08379000;
      W_f[10,1] := -0.16816668;
      W_f[10,2] := 0.01026458;
      W_f[10,3] := -0.05021837;
      W_f[10,4] := -0.08648673;
      W_f[10,5] := 0.05194992;
      W_f[10,6] := -0.04798879;
      W_f[10,7] := -0.00668964;
      W_f[10,8] := -0.01598040;
      W_f[10,9] := -0.19321908;
      W_f[10,10] := -0.00677647;
      W_f[10,11] := -0.11638412;
      W_f[10,12] := -0.05050007;
      W_f[10,13] := -0.05213704;
      W_f[10,14] := -0.18101706;
      W_f[10,15] := 0.02277401;
      W_f[10,16] := 0.02921080;
      W_f[10,17] := 0.00873813;
      W_f[10,18] := 0.06415650;
      W_f[10,19] := -0.08317487;
      W_f[10,20] := -0.02438755;
      W_f[10,21] := -0.16884466;
      W_f[10,22] := 0.27693939;
      W_f[10,23] := 0.00935439;
      W_f[10,24] := 1.43402386;
      W_f[10,25] := 1.74972332;
      W_f[10,26] := 0.01418469;
      W_f[10,27] := 0.14746916;
      W_f[10,28] := 0.17624062;
      W_f[10,29] := 0.38566202;
      W_f[10,30] := 0.24629667;
      W_f[10,31] := -0.06444994;
      W_f[10,32] := 0.02206947;
      W_f[10,33] := 0.01205150;
      W_f[10,34] := 0.64443576;
      W_f[10,35] := 0.17858964;
      W_f[10,36] := 0.02772049;
      W_f[10,37] := 0.09627288;
      W_f[10,38] := -0.00038884;
      W_f[10,39] := 0.09056027;
      W_f[11,0] := 0.04731990;
      W_f[11,1] := 0.07852971;
      W_f[11,2] := 0.04516530;
      W_f[11,3] := 0.08165582;
      W_f[11,4] := -0.00823189;
      W_f[11,5] := 0.03292342;
      W_f[11,6] := 0.08625521;
      W_f[11,7] := 0.03074309;
      W_f[11,8] := -0.06851767;
      W_f[11,9] := -0.02743477;
      W_f[11,10] := 0.00402056;
      W_f[11,11] := 0.01896705;
      W_f[11,12] := 0.02100093;
      W_f[11,13] := 0.04474377;
      W_f[11,14] := -0.03925331;
      W_f[11,15] := -0.01760299;
      W_f[11,16] := -0.05878574;
      W_f[11,17] := -0.00179996;
      W_f[11,18] := 0.01894562;
      W_f[11,19] := 0.01100245;
      W_f[11,20] := -0.08416440;
      W_f[11,21] := 0.08459154;
      W_f[11,22] := -0.07597429;
      W_f[11,23] := -0.02480526;
      W_f[11,24] := -0.30214685;
      W_f[11,25] := -0.06083889;
      W_f[11,26] := 0.05015881;
      W_f[11,27] := -0.01587165;
      W_f[11,28] := -0.00948480;
      W_f[11,29] := 0.16900283;
      W_f[11,30] := 0.01662034;
      W_f[11,31] := -0.04290604;
      W_f[11,32] := -0.15728204;
      W_f[11,33] := 0.18166886;
      W_f[11,34] := 0.06984576;
      W_f[11,35] := 0.02457202;
      W_f[11,36] := 0.02189556;
      W_f[11,37] := -0.02640078;
      W_f[11,38] := 0.00093580;
      W_f[11,39] := 0.04468563;
      W_f[12,0] := 0.13872766;
      W_f[12,1] := 0.36059234;
      W_f[12,2] := 0.18638378;
      W_f[12,3] := 0.38616773;
      W_f[12,4] := 0.18198954;
      W_f[12,5] := -0.01693199;
      W_f[12,6] := 0.51554531;
      W_f[12,7] := 0.66682684;
      W_f[12,8] := -0.49452236;
      W_f[12,9] := 0.56500375;
      W_f[12,10] := -0.31727192;
      W_f[12,11] := -0.16788831;
      W_f[12,12] := -0.09018624;
      W_f[12,13] := -0.02442008;
      W_f[12,14] := -0.06402968;
      W_f[12,15] := -0.11079653;
      W_f[12,16] := 0.23340648;
      W_f[12,17] := -0.03873094;
      W_f[12,18] := -0.35387737;
      W_f[12,19] := -0.13109617;
      W_f[12,20] := -0.02236723;
      W_f[12,21] := -0.25169286;
      W_f[12,22] := 0.04343348;
      W_f[12,23] := -0.14147434;
      W_f[12,24] := 0.09822226;
      W_f[12,25] := 0.07601354;
      W_f[12,26] := 0.13397673;
      W_f[12,27] := -0.16423117;
      W_f[12,28] := 0.20508496;
      W_f[12,29] := -0.19170563;
      W_f[12,30] := -0.21707255;
      W_f[12,31] := 0.19305049;
      W_f[12,32] := -0.00178745;
      W_f[12,33] := -0.02608595;
      W_f[12,34] := 0.07433556;
      W_f[12,35] := -0.07448775;
      W_f[12,36] := -0.12259015;
      W_f[12,37] := 0.05483592;
      W_f[12,38] := -0.02252366;
      W_f[12,39] := -0.13191852;
      W_f[13,0] := 0.05621623;
      W_f[13,1] := 0.02268710;
      W_f[13,2] := -0.02137025;
      W_f[13,3] := -0.03402603;
      W_f[13,4] := -0.00403033;
      W_f[13,5] := 0.05825109;
      W_f[13,6] := 0.02592259;
      W_f[13,7] := 0.01048357;
      W_f[13,8] := -0.00884827;
      W_f[13,9] := -0.07394934;
      W_f[13,10] := 0.01323845;
      W_f[13,11] := 0.11154817;
      W_f[13,12] := 0.19265266;
      W_f[13,13] := 0.09498972;
      W_f[13,14] := -0.01949506;
      W_f[13,15] := 0.01599856;
      W_f[13,16] := -0.04177938;
      W_f[13,17] := -0.01963896;
      W_f[13,18] := 0.06818765;
      W_f[13,19] := -0.10189550;
      W_f[13,20] := -0.00283599;
      W_f[13,21] := -0.02469871;
      W_f[13,22] := -0.04763987;
      W_f[13,23] := -0.05747910;
      W_f[13,24] := 0.62972993;
      W_f[13,25] := 0.50124347;
      W_f[13,26] := -0.15037754;
      W_f[13,27] := -0.02853806;
      W_f[13,28] := 0.03832513;
      W_f[13,29] := 0.01257216;
      W_f[13,30] := 0.03315365;
      W_f[13,31] := 0.00258718;
      W_f[13,32] := 0.23024213;
      W_f[13,33] := 0.01467210;
      W_f[13,34] := 0.52416134;
      W_f[13,35] := -0.07634575;
      W_f[13,36] := 0.00017335;
      W_f[13,37] := -0.06273333;
      W_f[13,38] := 0.01321615;
      W_f[13,39] := 0.01253699;
      W_f[14,0] := 0.05188091;
      W_f[14,1] := 0.09008571;
      W_f[14,2] := -0.06040832;
      W_f[14,3] := -0.15870132;
      W_f[14,4] := 0.01968341;
      W_f[14,5] := -0.02412392;
      W_f[14,6] := 0.00604502;
      W_f[14,7] := 0.00272764;
      W_f[14,8] := -0.02168215;
      W_f[14,9] := -0.08099962;
      W_f[14,10] := 0.01248098;
      W_f[14,11] := 0.04416423;
      W_f[14,12] := 0.01406407;
      W_f[14,13] := -0.03414071;
      W_f[14,14] := 0.00417258;
      W_f[14,15] := -0.15435918;
      W_f[14,16] := 0.11206103;
      W_f[14,17] := -0.05795342;
      W_f[14,18] := 0.20023122;
      W_f[14,19] := 0.25853318;
      W_f[14,20] := -0.04636193;
      W_f[14,21] := 0.05119645;
      W_f[14,22] := 0.01715696;
      W_f[14,23] := 0.00778349;
      W_f[14,24] := -0.25048414;
      W_f[14,25] := -0.59388351;
      W_f[14,26] := 0.12166926;
      W_f[14,27] := -0.01130306;
      W_f[14,28] := 0.02301564;
      W_f[14,29] := 0.03248704;
      W_f[14,30] := 0.04664331;
      W_f[14,31] := 0.05805317;
      W_f[14,32] := 0.02991675;
      W_f[14,33] := 0.12733400;
      W_f[14,34] := -0.05554454;
      W_f[14,35] := -0.04630656;
      W_f[14,36] := -0.04581423;
      W_f[14,37] := 0.15576649;
      W_f[14,38] := -0.03458373;
      W_f[14,39] := 0.07389181;
      W_f[15,0] := -0.02851857;
      W_f[15,1] := 0.12228543;
      W_f[15,2] := 0.04074666;
      W_f[15,3] := -0.16404167;
      W_f[15,4] := 0.03169363;
      W_f[15,5] := -0.04794145;
      W_f[15,6] := -0.02538486;
      W_f[15,7] := 0.09773283;
      W_f[15,8] := -0.00113020;
      W_f[15,9] := 0.00206907;
      W_f[15,10] := 0.00170394;
      W_f[15,11] := -0.18747102;
      W_f[15,12] := 0.13273963;
      W_f[15,13] := 0.00116777;
      W_f[15,14] := -0.01292728;
      W_f[15,15] := -0.05278755;
      W_f[15,16] := 0.02699348;
      W_f[15,17] := 0.06503567;
      W_f[15,18] := -0.08527236;
      W_f[15,19] := -0.36556801;
      W_f[15,20] := 0.04682306;
      W_f[15,21] := 0.18975946;
      W_f[15,22] := 0.58196318;
      W_f[15,23] := 0.01483520;
      W_f[15,24] := 1.57459116;
      W_f[15,25] := 1.53082824;
      W_f[15,26] := 0.08213925;
      W_f[15,27] := 0.17018035;
      W_f[15,28] := 0.16270036;
      W_f[15,29] := -1.25782382;
      W_f[15,30] := 0.78321606;
      W_f[15,31] := -0.03324566;
      W_f[15,32] := 0.06538258;
      W_f[15,33] := 0.22916409;
      W_f[15,34] := 1.10171151;
      W_f[15,35] := 0.06133924;
      W_f[15,36] := -0.06126631;
      W_f[15,37] := 0.05620775;
      W_f[15,38] := 0.02675290;
      W_f[15,39] := 0.08648319;
      W_g[0,0] := -0.03288272;
      W_g[0,1] := 0.06879283;
      W_g[0,2] := -0.02887416;
      W_g[0,3] := 0.02746971;
      W_g[0,4] := 0.04634671;
      W_g[0,5] := -0.01307166;
      W_g[0,6] := 0.04332437;
      W_g[0,7] := 0.02397616;
      W_g[0,8] := 0.02618686;
      W_g[0,9] := 0.02531774;
      W_g[0,10] := -0.00689762;
      W_g[0,11] := -0.03228850;
      W_g[0,12] := -0.04695914;
      W_g[0,13] := -0.00249899;
      W_g[0,14] := -0.06194285;
      W_g[0,15] := -0.01109950;
      W_g[0,16] := 0.00831518;
      W_g[0,17] := -0.11515938;
      W_g[0,18] := 0.00697446;
      W_g[0,19] := -0.06260984;
      W_g[0,20] := -0.06981920;
      W_g[0,21] := -0.10400263;
      W_g[0,22] := 0.00419812;
      W_g[0,23] := 0.02415262;
      W_g[0,24] := -0.13206881;
      W_g[0,25] := 0.14327736;
      W_g[0,26] := 0.07169567;
      W_g[0,27] := -0.13220897;
      W_g[0,28] := 0.07111509;
      W_g[0,29] := 0.00454173;
      W_g[0,30] := -0.00463334;
      W_g[0,31] := 0.00058220;
      W_g[0,32] := 0.00037708;
      W_g[0,33] := -0.00026135;
      W_g[0,34] := 0.22679581;
      W_g[0,35] := 0.00052285;
      W_g[0,36] := 0.00264373;
      W_g[0,37] := -0.02689169;
      W_g[0,38] := -0.00969260;
      W_g[0,39] := -0.03882377;
      W_g[1,0] := -0.05839003;
      W_g[1,1] := 0.42263713;
      W_g[1,2] := -0.04012571;
      W_g[1,3] := 0.01434622;
      W_g[1,4] := -0.05931747;
      W_g[1,5] := -0.09267445;
      W_g[1,6] := 0.09244086;
      W_g[1,7] := 0.00149189;
      W_g[1,8] := 0.01646185;
      W_g[1,9] := 0.00913838;
      W_g[1,10] := 0.01058344;
      W_g[1,11] := -0.03441796;
      W_g[1,12] := -0.02675500;
      W_g[1,13] := -0.01039137;
      W_g[1,14] := -0.02187960;
      W_g[1,15] := -0.03511444;
      W_g[1,16] := 0.06820389;
      W_g[1,17] := 0.00374079;
      W_g[1,18] := 0.09911744;
      W_g[1,19] := -0.02790303;
      W_g[1,20] := -0.21210110;
      W_g[1,21] := 0.14164248;
      W_g[1,22] := -0.04919457;
      W_g[1,23] := -0.10424531;
      W_g[1,24] := -0.25002548;
      W_g[1,25] := -0.41824010;
      W_g[1,26] := -0.05768240;
      W_g[1,27] := 0.16974758;
      W_g[1,28] := 0.08134635;
      W_g[1,29] := 0.01095367;
      W_g[1,30] := -0.10672898;
      W_g[1,31] := -0.03143495;
      W_g[1,32] := -0.05365749;
      W_g[1,33] := 0.00830225;
      W_g[1,34] := 0.00796971;
      W_g[1,35] := -0.11966703;
      W_g[1,36] := 0.10712396;
      W_g[1,37] := 0.04311150;
      W_g[1,38] := 0.02923429;
      W_g[1,39] := 0.00462070;
      W_g[2,0] := -0.01095263;
      W_g[2,1] := 0.07733528;
      W_g[2,2] := -0.00723971;
      W_g[2,3] := 0.00655987;
      W_g[2,4] := 0.05033382;
      W_g[2,5] := -0.05086170;
      W_g[2,6] := -0.00893102;
      W_g[2,7] := 0.00838173;
      W_g[2,8] := 0.01219127;
      W_g[2,9] := -0.00249959;
      W_g[2,10] := 0.01104422;
      W_g[2,11] := 0.08935806;
      W_g[2,12] := 0.05025892;
      W_g[2,13] := 0.01599896;
      W_g[2,14] := -0.14540766;
      W_g[2,15] := 0.03795051;
      W_g[2,16] := 0.00179014;
      W_g[2,17] := 0.12772407;
      W_g[2,18] := -0.09817299;
      W_g[2,19] := 0.13920712;
      W_g[2,20] := 0.00742573;
      W_g[2,21] := 0.00262788;
      W_g[2,22] := 0.01521684;
      W_g[2,23] := -0.00954701;
      W_g[2,24] := 0.62358665;
      W_g[2,25] := 0.38909104;
      W_g[2,26] := 0.02143394;
      W_g[2,27] := 0.01759339;
      W_g[2,28] := 0.06352523;
      W_g[2,29] := -0.04855579;
      W_g[2,30] := 0.02580756;
      W_g[2,31] := 0.00596368;
      W_g[2,32] := 0.01640637;
      W_g[2,33] := 0.02091035;
      W_g[2,34] := 0.49321541;
      W_g[2,35] := 0.03743263;
      W_g[2,36] := -0.01044649;
      W_g[2,37] := -0.00274277;
      W_g[2,38] := 0.00144159;
      W_g[2,39] := -0.59162003;
      W_g[3,0] := -0.02036412;
      W_g[3,1] := -0.14411704;
      W_g[3,2] := -0.02639455;
      W_g[3,3] := 0.02397250;
      W_g[3,4] := -0.16004682;
      W_g[3,5] := -0.00529983;
      W_g[3,6] := 0.13255818;
      W_g[3,7] := 0.02613736;
      W_g[3,8] := 0.01934580;
      W_g[3,9] := 0.02009285;
      W_g[3,10] := -0.06752108;
      W_g[3,11] := -0.04748070;
      W_g[3,12] := -0.05999199;
      W_g[3,13] := 0.00653862;
      W_g[3,14] := -0.03967655;
      W_g[3,15] := -0.03746946;
      W_g[3,16] := 0.02267453;
      W_g[3,17] := -0.07123119;
      W_g[3,18] := 0.03707521;
      W_g[3,19] := -0.06942015;
      W_g[3,20] := -0.10585976;
      W_g[3,21] := 0.07069318;
      W_g[3,22] := 0.04288564;
      W_g[3,23] := 0.09068061;
      W_g[3,24] := 0.25938836;
      W_g[3,25] := -0.00764711;
      W_g[3,26] := -0.00429336;
      W_g[3,27] := 0.10295356;
      W_g[3,28] := -0.12612087;
      W_g[3,29] := 0.00479916;
      W_g[3,30] := 0.15239407;
      W_g[3,31] := 0.05638619;
      W_g[3,32] := 0.05324322;
      W_g[3,33] := 0.03522293;
      W_g[3,34] := 0.02783547;
      W_g[3,35] := -0.00447224;
      W_g[3,36] := 0.34176287;
      W_g[3,37] := 0.15846112;
      W_g[3,38] := 0.02763572;
      W_g[3,39] := -0.00952189;
      W_g[4,0] := 0.05488009;
      W_g[4,1] := -0.00670369;
      W_g[4,2] := 0.04741509;
      W_g[4,3] := 0.00571730;
      W_g[4,4] := -0.06987662;
      W_g[4,5] := 0.01855648;
      W_g[4,6] := 0.09008339;
      W_g[4,7] := 0.00667926;
      W_g[4,8] := 0.00658040;
      W_g[4,9] := 0.00961057;
      W_g[4,10] := -0.04362585;
      W_g[4,11] := -0.03329441;
      W_g[4,12] := -0.01316141;
      W_g[4,13] := 0.14691545;
      W_g[4,14] := 0.00850634;
      W_g[4,15] := -0.05621828;
      W_g[4,16] := -0.05743054;
      W_g[4,17] := 0.13111739;
      W_g[4,18] := 0.00087735;
      W_g[4,19] := -0.02226411;
      W_g[4,20] := -0.11267117;
      W_g[4,21] := -0.02835003;
      W_g[4,22] := -0.02741843;
      W_g[4,23] := 0.13355793;
      W_g[4,24] := -0.16290458;
      W_g[4,25] := -0.17808466;
      W_g[4,26] := 0.02852475;
      W_g[4,27] := -0.02260069;
      W_g[4,28] := 0.03386381;
      W_g[4,29] := 0.04136939;
      W_g[4,30] := -0.02621254;
      W_g[4,31] := -0.02350034;
      W_g[4,32] := -0.02518253;
      W_g[4,33] := -0.02326495;
      W_g[4,34] := -0.32219490;
      W_g[4,35] := -0.05711325;
      W_g[4,36] := 0.05694984;
      W_g[4,37] := 0.00658011;
      W_g[4,38] := -0.06881828;
      W_g[4,39] := -0.02566535;
      W_g[5,0] := -0.12075401;
      W_g[5,1] := 0.02553332;
      W_g[5,2] := -0.12287396;
      W_g[5,3] := 0.12021825;
      W_g[5,4] := -0.07048963;
      W_g[5,5] := -0.14113422;
      W_g[5,6] := 0.05872258;
      W_g[5,7] := 0.12207281;
      W_g[5,8] := 0.11423667;
      W_g[5,9] := 0.12041245;
      W_g[5,10] := 0.01521803;
      W_g[5,11] := -0.01810576;
      W_g[5,12] := -0.00813478;
      W_g[5,13] := -0.08835436;
      W_g[5,14] := 0.09394597;
      W_g[5,15] := -0.04471128;
      W_g[5,16] := -0.06250727;
      W_g[5,17] := 0.06817933;
      W_g[5,18] := -0.01152834;
      W_g[5,19] := -0.00579273;
      W_g[5,20] := -0.08372810;
      W_g[5,21] := -0.06996331;
      W_g[5,22] := 0.01203206;
      W_g[5,23] := 0.00779026;
      W_g[5,24] := 0.08353818;
      W_g[5,25] := -0.25279960;
      W_g[5,26] := 0.05011104;
      W_g[5,27] := -0.10751224;
      W_g[5,28] := -0.07444005;
      W_g[5,29] := -0.02102967;
      W_g[5,30] := 0.00832473;
      W_g[5,31] := 0.01262962;
      W_g[5,32] := -0.01239251;
      W_g[5,33] := 0.00079978;
      W_g[5,34] := 0.07374854;
      W_g[5,35] := -0.04611919;
      W_g[5,36] := -0.01176891;
      W_g[5,37] := 0.02829348;
      W_g[5,38] := 0.00393110;
      W_g[5,39] := 0.07769092;
      W_g[6,0] := -0.05814515;
      W_g[6,1] := -0.04702876;
      W_g[6,2] := -0.06337287;
      W_g[6,3] := 0.03413104;
      W_g[6,4] := 0.06652597;
      W_g[6,5] := -0.05150583;
      W_g[6,6] := -0.01204906;
      W_g[6,7] := 0.03913860;
      W_g[6,8] := 0.03228532;
      W_g[6,9] := 0.03164063;
      W_g[6,10] := 0.01173771;
      W_g[6,11] := -0.01391642;
      W_g[6,12] := -0.03429415;
      W_g[6,13] := -0.04339701;
      W_g[6,14] := 0.06324015;
      W_g[6,15] := -0.00640369;
      W_g[6,16] := 0.18601589;
      W_g[6,17] := -0.00700807;
      W_g[6,18] := 0.00076136;
      W_g[6,19] := -0.05252279;
      W_g[6,20] := 0.04849189;
      W_g[6,21] := 0.02619516;
      W_g[6,22] := -0.00269682;
      W_g[6,23] := -0.02741523;
      W_g[6,24] := 0.05987318;
      W_g[6,25] := 0.04793175;
      W_g[6,26] := -0.02643443;
      W_g[6,27] := 0.04390920;
      W_g[6,28] := 0.03213611;
      W_g[6,29] := 0.01188661;
      W_g[6,30] := -0.01111693;
      W_g[6,31] := -0.00252879;
      W_g[6,32] := -0.00546005;
      W_g[6,33] := -0.00067087;
      W_g[6,34] := 0.17834580;
      W_g[6,35] := 0.00388802;
      W_g[6,36] := -0.02650490;
      W_g[6,37] := 0.01564691;
      W_g[6,38] := -0.30253130;
      W_g[6,39] := -0.15068348;
      W_g[7,0] := -0.10275671;
      W_g[7,1] := -0.24009611;
      W_g[7,2] := -0.11088440;
      W_g[7,3] := -0.01006387;
      W_g[7,4] := -0.03458254;
      W_g[7,5] := 0.23932587;
      W_g[7,6] := 0.40470347;
      W_g[7,7] := -0.00585874;
      W_g[7,8] := -0.01916949;
      W_g[7,9] := -0.00627702;
      W_g[7,10] := -0.27911651;
      W_g[7,11] := 0.01163200;
      W_g[7,12] := 0.01657399;
      W_g[7,13] := -0.10315786;
      W_g[7,14] := 0.03309733;
      W_g[7,15] := 0.00751682;
      W_g[7,16] := -0.02915282;
      W_g[7,17] := 0.03935070;
      W_g[7,18] := -0.12759872;
      W_g[7,19] := 0.04157587;
      W_g[7,20] := -0.30659992;
      W_g[7,21] := 0.09425942;
      W_g[7,22] := -0.00641260;
      W_g[7,23] := -0.09050559;
      W_g[7,24] := 0.01530947;
      W_g[7,25] := -0.15979554;
      W_g[7,26] := -0.00322467;
      W_g[7,27] := 0.04318399;
      W_g[7,28] := 0.14858317;
      W_g[7,29] := 0.04615099;
      W_g[7,30] := 0.00307166;
      W_g[7,31] := 0.04133423;
      W_g[7,32] := 0.00097957;
      W_g[7,33] := 0.02065461;
      W_g[7,34] := 0.04547579;
      W_g[7,35] := -0.00785838;
      W_g[7,36] := -0.20765284;
      W_g[7,37] := 0.00956008;
      W_g[7,38] := 0.00075457;
      W_g[7,39] := 0.02893667;
      W_g[8,0] := -0.08692090;
      W_g[8,1] := 0.08997668;
      W_g[8,2] := -0.09005233;
      W_g[8,3] := -0.01292246;
      W_g[8,4] := 0.10805142;
      W_g[8,5] := 0.14603932;
      W_g[8,6] := -0.02134521;
      W_g[8,7] := -0.01256517;
      W_g[8,8] := -0.01110261;
      W_g[8,9] := -0.01626757;
      W_g[8,10] := 0.05898210;
      W_g[8,11] := -0.11047587;
      W_g[8,12] := -0.09589648;
      W_g[8,13] := -0.02350931;
      W_g[8,14] := 0.02544193;
      W_g[8,15] := -0.13092923;
      W_g[8,16] := 0.10931896;
      W_g[8,17] := 0.12825854;
      W_g[8,18] := 0.12620327;
      W_g[8,19] := -0.12419707;
      W_g[8,20] := 0.03848997;
      W_g[8,21] := -0.06537959;
      W_g[8,22] := 0.00064196;
      W_g[8,23] := -0.03796872;
      W_g[8,24] := -0.04377631;
      W_g[8,25] := -0.30099538;
      W_g[8,26] := 0.02286426;
      W_g[8,27] := -0.06000912;
      W_g[8,28] := 0.03258165;
      W_g[8,29] := -0.02475458;
      W_g[8,30] := -0.00219198;
      W_g[8,31] := -0.00292637;
      W_g[8,32] := 0.00115337;
      W_g[8,33] := 0.00390999;
      W_g[8,34] := -0.04075257;
      W_g[8,35] := -0.02803931;
      W_g[8,36] := 0.02655412;
      W_g[8,37] := 0.02139529;
      W_g[8,38] := 0.04244001;
      W_g[8,39] := 0.03061243;
      W_g[9,0] := -0.22739998;
      W_g[9,1] := -0.12028531;
      W_g[9,2] := -0.22718781;
      W_g[9,3] := -0.18262891;
      W_g[9,4] := -0.01637146;
      W_g[9,5] := -0.23831372;
      W_g[9,6] := 0.00297750;
      W_g[9,7] := -0.17095226;
      W_g[9,8] := -0.18344788;
      W_g[9,9] := -0.18747538;
      W_g[9,10] := -0.31918642;
      W_g[9,11] := -0.01426092;
      W_g[9,12] := -0.00200754;
      W_g[9,13] := 0.00886641;
      W_g[9,14] := -0.01517866;
      W_g[9,15] := -0.00491453;
      W_g[9,16] := 0.03928856;
      W_g[9,17] := 0.05202412;
      W_g[9,18] := -0.04777612;
      W_g[9,19] := 0.00385900;
      W_g[9,20] := 0.04262874;
      W_g[9,21] := -0.05054115;
      W_g[9,22] := -0.04248414;
      W_g[9,23] := -0.00319653;
      W_g[9,24] := -0.31163967;
      W_g[9,25] := -0.09675232;
      W_g[9,26] := -0.01050112;
      W_g[9,27] := -0.05346175;
      W_g[9,28] := -0.06083639;
      W_g[9,29] := 0.12653194;
      W_g[9,30] := -0.05285788;
      W_g[9,31] := -0.01213977;
      W_g[9,32] := -0.04765768;
      W_g[9,33] := -0.05291987;
      W_g[9,34] := -0.29435629;
      W_g[9,35] := -0.06011635;
      W_g[9,36] := -0.05353123;
      W_g[9,37] := 0.00832208;
      W_g[9,38] := 0.00973149;
      W_g[9,39] := -0.01172841;
      W_g[10,0] := 0.03514115;
      W_g[10,1] := 0.11389200;
      W_g[10,2] := 0.03716018;
      W_g[10,3] := -0.01071796;
      W_g[10,4] := -0.30562735;
      W_g[10,5] := 0.01998116;
      W_g[10,6] := 0.14969940;
      W_g[10,7] := -0.02109131;
      W_g[10,8] := -0.01540629;
      W_g[10,9] := -0.00982767;
      W_g[10,10] := -0.09813343;
      W_g[10,11] := -0.09390774;
      W_g[10,12] := -0.09303362;
      W_g[10,13] := -0.00659447;
      W_g[10,14] := -0.08698983;
      W_g[10,15] := -0.09059508;
      W_g[10,16] := -0.01796200;
      W_g[10,17] := -0.02903299;
      W_g[10,18] := 0.13222115;
      W_g[10,19] := -0.13716845;
      W_g[10,20] := -0.15225135;
      W_g[10,21] := 0.03876633;
      W_g[10,22] := 0.04551086;
      W_g[10,23] := 0.02596399;
      W_g[10,24] := 0.15688412;
      W_g[10,25] := 0.16100781;
      W_g[10,26] := 0.01107862;
      W_g[10,27] := -0.07539947;
      W_g[10,28] := -0.25086227;
      W_g[10,29] := -0.12395287;
      W_g[10,30] := 0.05308864;
      W_g[10,31] := 0.06245262;
      W_g[10,32] := 0.03307296;
      W_g[10,33] := 0.04681247;
      W_g[10,34] := 0.23864536;
      W_g[10,35] := 0.01017979;
      W_g[10,36] := -0.34682098;
      W_g[10,37] := 0.01139926;
      W_g[10,38] := -0.06640822;
      W_g[10,39] := -0.07425395;
      W_g[11,0] := -0.20998149;
      W_g[11,1] := 0.05767135;
      W_g[11,2] := -0.23170957;
      W_g[11,3] := 0.02501687;
      W_g[11,4] := 0.02252023;
      W_g[11,5] := 0.03745016;
      W_g[11,6] := 0.00724144;
      W_g[11,7] := 0.03957897;
      W_g[11,8] := 0.02575030;
      W_g[11,9] := 0.03189280;
      W_g[11,10] := 0.05883392;
      W_g[11,11] := 0.02762088;
      W_g[11,12] := 0.01796787;
      W_g[11,13] := 0.28403825;
      W_g[11,14] := 0.06086168;
      W_g[11,15] := 0.02774396;
      W_g[11,16] := 0.03697228;
      W_g[11,17] := -0.07755503;
      W_g[11,18] := -0.01424372;
      W_g[11,19] := 0.01996346;
      W_g[11,20] := 0.13414641;
      W_g[11,21] := 0.12937231;
      W_g[11,22] := -0.01583524;
      W_g[11,23] := 0.26789898;
      W_g[11,24] := 0.32321972;
      W_g[11,25] := 0.31935814;
      W_g[11,26] := -0.05019195;
      W_g[11,27] := 0.23280673;
      W_g[11,28] := 0.09163668;
      W_g[11,29] := -0.01618287;
      W_g[11,30] := -0.00085428;
      W_g[11,31] := -0.01937335;
      W_g[11,32] := 0.01763184;
      W_g[11,33] := -0.00380951;
      W_g[11,34] := 0.07600094;
      W_g[11,35] := 0.09330983;
      W_g[11,36] := -0.07791516;
      W_g[11,37] := 0.01969607;
      W_g[11,38] := 0.04727592;
      W_g[11,39] := 0.04515434;
      W_g[12,0] := -0.05593645;
      W_g[12,1] := -0.04389839;
      W_g[12,2] := -0.05817224;
      W_g[12,3] := 0.04144620;
      W_g[12,4] := -0.02310878;
      W_g[12,5] := 0.04852642;
      W_g[12,6] := -0.08700307;
      W_g[12,7] := 0.03355748;
      W_g[12,8] := 0.03699837;
      W_g[12,9] := 0.03886550;
      W_g[12,10] := 0.10981326;
      W_g[12,11] := -0.09832872;
      W_g[12,12] := -0.09303018;
      W_g[12,13] := -0.04333979;
      W_g[12,14] := -0.11123282;
      W_g[12,15] := -0.09018178;
      W_g[12,16] := -0.00510190;
      W_g[12,17] := -0.01573442;
      W_g[12,18] := -0.70857680;
      W_g[12,19] := -0.04782427;
      W_g[12,20] := 0.08851119;
      W_g[12,21] := 0.02074307;
      W_g[12,22] := -0.01258304;
      W_g[12,23] := -0.00788189;
      W_g[12,24] := -0.11268676;
      W_g[12,25] := -0.11553165;
      W_g[12,26] := -0.01619464;
      W_g[12,27] := 0.04248659;
      W_g[12,28] := -0.07553757;
      W_g[12,29] := 0.02218230;
      W_g[12,30] := -0.02093006;
      W_g[12,31] := -0.01882189;
      W_g[12,32] := -0.01577668;
      W_g[12,33] := -0.00407436;
      W_g[12,34] := -0.14571649;
      W_g[12,35] := -0.03193094;
      W_g[12,36] := 0.03408330;
      W_g[12,37] := -0.00389380;
      W_g[12,38] := 0.02884003;
      W_g[12,39] := -0.03945985;
      W_g[13,0] := 0.04027861;
      W_g[13,1] := -0.07311103;
      W_g[13,2] := 0.04157875;
      W_g[13,3] := 0.01889602;
      W_g[13,4] := -0.11995003;
      W_g[13,5] := -0.01993360;
      W_g[13,6] := 0.03187145;
      W_g[13,7] := 0.01748616;
      W_g[13,8] := 0.01463885;
      W_g[13,9] := 0.02840340;
      W_g[13,10] := -0.02596055;
      W_g[13,11] := 0.02591357;
      W_g[13,12] := 0.02623175;
      W_g[13,13] := -0.00677697;
      W_g[13,14] := -0.00711890;
      W_g[13,15] := 0.05769501;
      W_g[13,16] := 0.30919826;
      W_g[13,17] := 0.02394222;
      W_g[13,18] := -0.03814467;
      W_g[13,19] := 0.01873361;
      W_g[13,20] := -0.05235977;
      W_g[13,21] := -0.04417822;
      W_g[13,22] := -0.01057172;
      W_g[13,23] := 0.04463968;
      W_g[13,24] := 0.05050629;
      W_g[13,25] := -0.15972561;
      W_g[13,26] := 0.02774286;
      W_g[13,27] := -0.08080220;
      W_g[13,28] := -0.09933943;
      W_g[13,29] := 0.03062030;
      W_g[13,30] := -0.00385746;
      W_g[13,31] := 0.01280402;
      W_g[13,32] := -0.00358380;
      W_g[13,33] := -0.00492619;
      W_g[13,34] := 0.04224548;
      W_g[13,35] := -0.00044207;
      W_g[13,36] := -0.04630874;
      W_g[13,37] := -0.03753048;
      W_g[13,38] := 0.09008476;
      W_g[13,39] := 0.02002463;
      W_g[14,0] := 0.06269035;
      W_g[14,1] := 0.16204342;
      W_g[14,2] := 0.07219669;
      W_g[14,3] := -0.04503014;
      W_g[14,4] := -0.00555789;
      W_g[14,5] := 0.01761685;
      W_g[14,6] := -0.03159415;
      W_g[14,7] := -0.05064076;
      W_g[14,8] := -0.04640801;
      W_g[14,9] := -0.06009993;
      W_g[14,10] := 0.00660122;
      W_g[14,11] := -0.03258261;
      W_g[14,12] := -0.03601762;
      W_g[14,13] := 0.03453247;
      W_g[14,14] := 0.12738688;
      W_g[14,15] := -0.01328611;
      W_g[14,16] := 0.01626320;
      W_g[14,17] := -0.04504346;
      W_g[14,18] := -0.15708502;
      W_g[14,19] := 0.00090277;
      W_g[14,20] := -0.04051626;
      W_g[14,21] := -0.04047279;
      W_g[14,22] := 0.00840584;
      W_g[14,23] := -0.01122396;
      W_g[14,24] := 0.06744422;
      W_g[14,25] := 0.49537152;
      W_g[14,26] := 0.07856539;
      W_g[14,27] := -0.03960157;
      W_g[14,28] := 0.03958257;
      W_g[14,29] := -0.04088740;
      W_g[14,30] := 0.02040378;
      W_g[14,31] := 0.01003806;
      W_g[14,32] := 0.02256208;
      W_g[14,33] := 0.02816826;
      W_g[14,34] := 0.15040024;
      W_g[14,35] := 0.01636149;
      W_g[14,36] := 0.04578492;
      W_g[14,37] := -0.03131405;
      W_g[14,38] := -0.05991198;
      W_g[14,39] := 0.01529666;
      W_g[15,0] := 0.11327556;
      W_g[15,1] := -0.17608264;
      W_g[15,2] := 0.09651362;
      W_g[15,3] := 0.02762307;
      W_g[15,4] := 0.26826185;
      W_g[15,5] := -0.27072880;
      W_g[15,6] := 0.04821723;
      W_g[15,7] := 0.03941977;
      W_g[15,8] := 0.02793526;
      W_g[15,9] := 0.03359088;
      W_g[15,10] := -0.12275329;
      W_g[15,11] := -0.16014972;
      W_g[15,12] := -0.16786559;
      W_g[15,13] := 0.09324758;
      W_g[15,14] := -0.00898216;
      W_g[15,15] := -0.16123867;
      W_g[15,16] := 0.02021289;
      W_g[15,17] := -0.01648896;
      W_g[15,18] := -0.00597759;
      W_g[15,19] := -0.16053081;
      W_g[15,20] := 0.04093139;
      W_g[15,21] := 0.06445049;
      W_g[15,22] := 0.04804592;
      W_g[15,23] := 0.06335551;
      W_g[15,24] := 0.06702932;
      W_g[15,25] := 0.00881007;
      W_g[15,26] := 0.00152106;
      W_g[15,27] := 0.07652006;
      W_g[15,28] := 0.30222309;
      W_g[15,29] := -0.08014103;
      W_g[15,30] := 0.06666484;
      W_g[15,31] := 0.00829429;
      W_g[15,32] := 0.10078011;
      W_g[15,33] := 0.06581395;
      W_g[15,34] := 0.08893893;
      W_g[15,35] := 0.15266605;
      W_g[15,36] := -0.17053175;
      W_g[15,37] := -0.07062726;
      W_g[15,38] := 0.07771596;
      W_g[15,39] := 0.04211254;
      W_o[0,0] := 0.12198126;
      W_o[0,1] := 0.14187956;
      W_o[0,2] := -0.01325197;
      W_o[0,3] := -0.07755501;
      W_o[0,4] := -0.21710020;
      W_o[0,5] := 0.13306709;
      W_o[0,6] := -0.10178271;
      W_o[0,7] := -0.14437862;
      W_o[0,8] := 0.02041168;
      W_o[0,9] := 0.04337119;
      W_o[0,10] := 0.22460431;
      W_o[0,11] := -0.27840534;
      W_o[0,12] := 0.35424832;
      W_o[0,13] := 0.20462060;
      W_o[0,14] := -0.34063420;
      W_o[0,15] := 0.18119343;
      W_o[0,16] := -0.08057553;
      W_o[0,17] := -0.48889911;
      W_o[0,18] := 0.81621987;
      W_o[0,19] := 0.08914678;
      W_o[0,20] := 0.22458921;
      W_o[0,21] := 0.74807531;
      W_o[0,22] := 0.98743701;
      W_o[0,23] := -0.22151884;
      W_o[0,24] := 1.91302598;
      W_o[0,25] := 2.06443334;
      W_o[0,26] := -0.67687452;
      W_o[0,27] := -0.00083833;
      W_o[0,28] := -0.11211787;
      W_o[0,29] := -0.28486133;
      W_o[0,30] := 0.70833492;
      W_o[0,31] := 0.04462677;
      W_o[0,32] := 0.38353100;
      W_o[0,33] := 0.09996076;
      W_o[0,34] := 1.72650719;
      W_o[0,35] := 0.41856179;
      W_o[0,36] := 0.03231431;
      W_o[0,37] := 0.25164288;
      W_o[0,38] := 0.06612357;
      W_o[0,39] := -0.00002071;
      W_o[1,0] := -0.03910590;
      W_o[1,1] := 0.27588379;
      W_o[1,2] := 0.10975786;
      W_o[1,3] := -0.09756759;
      W_o[1,4] := -0.59621233;
      W_o[1,5] := -0.42031246;
      W_o[1,6] := -0.09698014;
      W_o[1,7] := 0.15754665;
      W_o[1,8] := -0.00284551;
      W_o[1,9] := 0.02527599;
      W_o[1,10] := -0.01773636;
      W_o[1,11] := -0.30956084;
      W_o[1,12] := 0.23456147;
      W_o[1,13] := 0.24187891;
      W_o[1,14] := 0.16774826;
      W_o[1,15] := 0.13618931;
      W_o[1,16] := -0.05666412;
      W_o[1,17] := -0.01989032;
      W_o[1,18] := -0.31193376;
      W_o[1,19] := -0.24264094;
      W_o[1,20] := -0.49747720;
      W_o[1,21] := 0.33921909;
      W_o[1,22] := -0.08854222;
      W_o[1,23] := 0.46807775;
      W_o[1,24] := -0.29946747;
      W_o[1,25] := -0.03667294;
      W_o[1,26] := 0.20074379;
      W_o[1,27] := 0.39029807;
      W_o[1,28] := -0.37250715;
      W_o[1,29] := -0.00592554;
      W_o[1,30] := -0.22806711;
      W_o[1,31] := -0.08731094;
      W_o[1,32] := -0.04087760;
      W_o[1,33] := 0.00680849;
      W_o[1,34] := -0.19797693;
      W_o[1,35] := -0.33509916;
      W_o[1,36] := 0.24450488;
      W_o[1,37] := -0.10827561;
      W_o[1,38] := 0.90532941;
      W_o[1,39] := 0.24546179;
      W_o[2,0] := -0.00616825;
      W_o[2,1] := 0.13651501;
      W_o[2,2] := -0.09869462;
      W_o[2,3] := -0.07334173;
      W_o[2,4] := -0.02211194;
      W_o[2,5] := 0.05619258;
      W_o[2,6] := 0.10801718;
      W_o[2,7] := 0.14577843;
      W_o[2,8] := 0.09542450;
      W_o[2,9] := 0.04769905;
      W_o[2,10] := 0.04124768;
      W_o[2,11] := -0.33887896;
      W_o[2,12] := 0.43093050;
      W_o[2,13] := 0.04022788;
      W_o[2,14] := 0.01084119;
      W_o[2,15] := 0.23125160;
      W_o[2,16] := 0.00388798;
      W_o[2,17] := -0.03658837;
      W_o[2,18] := -0.47197291;
      W_o[2,19] := 0.30483419;
      W_o[2,20] := -0.05675438;
      W_o[2,21] := -0.20610483;
      W_o[2,22] := -0.15346101;
      W_o[2,23] := -0.01675959;
      W_o[2,24] := -0.10398360;
      W_o[2,25] := 0.05681018;
      W_o[2,26] := -0.06196046;
      W_o[2,27] := 0.19941610;
      W_o[2,28] := 0.04805862;
      W_o[2,29] := 0.23355408;
      W_o[2,30] := -0.05858275;
      W_o[2,31] := -0.03168040;
      W_o[2,32] := -0.18688639;
      W_o[2,33] := 0.00733624;
      W_o[2,34] := 0.03196214;
      W_o[2,35] := -0.02429556;
      W_o[2,36] := -0.04773033;
      W_o[2,37] := -0.08787826;
      W_o[2,38] := 0.01416256;
      W_o[2,39] := 0.77567047;
      W_o[3,0] := 0.21000762;
      W_o[3,1] := 0.56502008;
      W_o[3,2] := 0.01591207;
      W_o[3,3] := -0.11321840;
      W_o[3,4] := 0.23269446;
      W_o[3,5] := 0.09338996;
      W_o[3,6] := 0.12135104;
      W_o[3,7] := 0.30009910;
      W_o[3,8] := 0.28139746;
      W_o[3,9] := -0.11283773;
      W_o[3,10] := -0.12950897;
      W_o[3,11] := -0.16686824;
      W_o[3,12] := 0.02030786;
      W_o[3,13] := 0.21336913;
      W_o[3,14] := -0.06828818;
      W_o[3,15] := -0.10707476;
      W_o[3,16] := 0.01645426;
      W_o[3,17] := -0.08346992;
      W_o[3,18] := 0.58030689;
      W_o[3,19] := 0.02444929;
      W_o[3,20] := -0.22163415;
      W_o[3,21] := 0.61291105;
      W_o[3,22] := -0.28959793;
      W_o[3,23] := -0.06618109;
      W_o[3,24] := 0.31345260;
      W_o[3,25] := 0.13633017;
      W_o[3,26] := -0.08859906;
      W_o[3,27] := -0.25854555;
      W_o[3,28] := -0.18073046;
      W_o[3,29] := -0.06065677;
      W_o[3,30] := -0.42247161;
      W_o[3,31] := 0.19295032;
      W_o[3,32] := -0.42941913;
      W_o[3,33] := 0.22519505;
      W_o[3,34] := -0.16697113;
      W_o[3,35] := -0.12213719;
      W_o[3,36] := 0.07402483;
      W_o[3,37] := -0.18623771;
      W_o[3,38] := -0.06633836;
      W_o[3,39] := -0.00843535;
      W_o[4,0] := -0.08241624;
      W_o[4,1] := -0.15822247;
      W_o[4,2] := -0.10238844;
      W_o[4,3] := -0.03743736;
      W_o[4,4] := 0.04915955;
      W_o[4,5] := 0.13049453;
      W_o[4,6] := 0.17377743;
      W_o[4,7] := -0.06675444;
      W_o[4,8] := -0.03882149;
      W_o[4,9] := 0.06404497;
      W_o[4,10] := 0.00192631;
      W_o[4,11] := -0.45325428;
      W_o[4,12] := 0.25542077;
      W_o[4,13] := -0.36887005;
      W_o[4,14] := -0.18856272;
      W_o[4,15] := -0.13098666;
      W_o[4,16] := -0.22178020;
      W_o[4,17] := -0.29496050;
      W_o[4,18] := -0.00731075;
      W_o[4,19] := -0.09241781;
      W_o[4,20] := -0.26850891;
      W_o[4,21] := -0.20041393;
      W_o[4,22] := -0.53797185;
      W_o[4,23] := 0.50577527;
      W_o[4,24] := 0.98513478;
      W_o[4,25] := 1.10475135;
      W_o[4,26] := 0.09366516;
      W_o[4,27] := 0.19566087;
      W_o[4,28] := -0.13328505;
      W_o[4,29] := 0.94272023;
      W_o[4,30] := -0.46258932;
      W_o[4,31] := -0.09195930;
      W_o[4,32] := -0.36374816;
      W_o[4,33] := -0.29488632;
      W_o[4,34] := 0.08194333;
      W_o[4,35] := -0.11618637;
      W_o[4,36] := -0.10650394;
      W_o[4,37] := -0.00409420;
      W_o[4,38] := 0.08796127;
      W_o[4,39] := 0.13779099;
      W_o[5,0] := 0.00298015;
      W_o[5,1] := 0.14726847;
      W_o[5,2] := -0.24877922;
      W_o[5,3] := 0.03818390;
      W_o[5,4] := 0.25190380;
      W_o[5,5] := 0.09698023;
      W_o[5,6] := 0.03788623;
      W_o[5,7] := -0.32500836;
      W_o[5,8] := -0.47933936;
      W_o[5,9] := -0.17586684;
      W_o[5,10] := 0.30961692;
      W_o[5,11] := -0.56706995;
      W_o[5,12] := -0.13458350;
      W_o[5,13] := 0.30265138;
      W_o[5,14] := 0.28882200;
      W_o[5,15] := -0.02685931;
      W_o[5,16] := 0.24619135;
      W_o[5,17] := 0.35931662;
      W_o[5,18] := 0.34230548;
      W_o[5,19] := 0.21314520;
      W_o[5,20] := 0.00126743;
      W_o[5,21] := 0.08332776;
      W_o[5,22] := 0.14433613;
      W_o[5,23] := -0.15501527;
      W_o[5,24] := 1.35550761;
      W_o[5,25] := 1.45758998;
      W_o[5,26] := -0.42872009;
      W_o[5,27] := 0.11975341;
      W_o[5,28] := 0.12516311;
      W_o[5,29] := -0.25945181;
      W_o[5,30] := 0.03064806;
      W_o[5,31] := -0.06416538;
      W_o[5,32] := 0.31372464;
      W_o[5,33] := 0.25143003;
      W_o[5,34] := 1.32014525;
      W_o[5,35] := 0.40504000;
      W_o[5,36] := 0.00424331;
      W_o[5,37] := 0.38437104;
      W_o[5,38] := 2.31802607;
      W_o[5,39] := 0.42288464;
      W_o[6,0] := 0.16465783;
      W_o[6,1] := -0.00748923;
      W_o[6,2] := -0.15153547;
      W_o[6,3] := -0.01711627;
      W_o[6,4] := -0.16756265;
      W_o[6,5] := 0.34808365;
      W_o[6,6] := 0.00590673;
      W_o[6,7] := -0.27918947;
      W_o[6,8] := 0.17359419;
      W_o[6,9] := 0.49527067;
      W_o[6,10] := -0.00244592;
      W_o[6,11] := -0.14789435;
      W_o[6,12] := 0.29600164;
      W_o[6,13] := -0.48868799;
      W_o[6,14] := -0.21440262;
      W_o[6,15] := -0.28105071;
      W_o[6,16] := 0.27140900;
      W_o[6,17] := -0.17575939;
      W_o[6,18] := 0.43315357;
      W_o[6,19] := 0.25442523;
      W_o[6,20] := 0.02021864;
      W_o[6,21] := 0.36727905;
      W_o[6,22] := 0.55856705;
      W_o[6,23] := 0.36519867;
      W_o[6,24] := 1.27994967;
      W_o[6,25] := 1.31188405;
      W_o[6,26] := 0.44206235;
      W_o[6,27] := 0.09447443;
      W_o[6,28] := 0.11994729;
      W_o[6,29] := -0.26271847;
      W_o[6,30] := 0.48323816;
      W_o[6,31] := -0.07709061;
      W_o[6,32] := 0.14690454;
      W_o[6,33] := 0.00670793;
      W_o[6,34] := 1.35142434;
      W_o[6,35] := 0.04027350;
      W_o[6,36] := 0.06238577;
      W_o[6,37] := 0.32636163;
      W_o[6,38] := -0.25480887;
      W_o[6,39] := 1.13409173;
      W_o[7,0] := 0.07718845;
      W_o[7,1] := 0.20402764;
      W_o[7,2] := 0.06463404;
      W_o[7,3] := 0.02887609;
      W_o[7,4] := -0.05794537;
      W_o[7,5] := 0.19518182;
      W_o[7,6] := 1.15763307;
      W_o[7,7] := 0.05626965;
      W_o[7,8] := 0.02816673;
      W_o[7,9] := 0.21392144;
      W_o[7,10] := -0.00420654;
      W_o[7,11] := -0.07277058;
      W_o[7,12] := 0.01088039;
      W_o[7,13] := 0.02142877;
      W_o[7,14] := -0.03849939;
      W_o[7,15] := -0.00698312;
      W_o[7,16] := 0.03512425;
      W_o[7,17] := -0.04141184;
      W_o[7,18] := 0.92844951;
      W_o[7,19] := -0.03062460;
      W_o[7,20] := -0.92607880;
      W_o[7,21] := 0.08325810;
      W_o[7,22] := 0.01044585;
      W_o[7,23] := -0.09986506;
      W_o[7,24] := -0.72718900;
      W_o[7,25] := -0.64502668;
      W_o[7,26] := -0.01259396;
      W_o[7,27] := -0.03038958;
      W_o[7,28] := -0.07504132;
      W_o[7,29] := 0.10145313;
      W_o[7,30] := -0.00330979;
      W_o[7,31] := 0.02509710;
      W_o[7,32] := -0.08854815;
      W_o[7,33] := -0.00711671;
      W_o[7,34] := -0.57390833;
      W_o[7,35] := -0.28441957;
      W_o[7,36] := 0.17795981;
      W_o[7,37] := -0.04241760;
      W_o[7,38] := -0.02305064;
      W_o[7,39] := -0.03192819;
      W_o[8,0] := -0.70497924;
      W_o[8,1] := -0.09449001;
      W_o[8,2] := -0.32517871;
      W_o[8,3] := 0.07309260;
      W_o[8,4] := -0.19864593;
      W_o[8,5] := 0.73818827;
      W_o[8,6] := -0.25948462;
      W_o[8,7] := 0.16984719;
      W_o[8,8] := -0.11935160;
      W_o[8,9] := 0.33245274;
      W_o[8,10] := 0.01087483;
      W_o[8,11] := -1.00101554;
      W_o[8,12] := -0.22074799;
      W_o[8,13] := 0.33614793;
      W_o[8,14] := -0.08536271;
      W_o[8,15] := -0.76774424;
      W_o[8,16] := 0.77750182;
      W_o[8,17] := 0.66594493;
      W_o[8,18] := 0.34620020;
      W_o[8,19] := 0.05137411;
      W_o[8,20] := -0.50151187;
      W_o[8,21] := -0.05596393;
      W_o[8,22] := 0.07904742;
      W_o[8,23] := -0.21896000;
      W_o[8,24] := 0.38224426;
      W_o[8,25] := 0.27276328;
      W_o[8,26] := 0.18764874;
      W_o[8,27] := -0.09256534;
      W_o[8,28] := -0.30482879;
      W_o[8,29] := 0.34679717;
      W_o[8,30] := -0.25258273;
      W_o[8,31] := 0.11198672;
      W_o[8,32] := 0.27686685;
      W_o[8,33] := 0.17793770;
      W_o[8,34] := 0.20446144;
      W_o[8,35] := -0.07079878;
      W_o[8,36] := -0.06305701;
      W_o[8,37] := 0.06945456;
      W_o[8,38] := 0.34880602;
      W_o[8,39] := -0.30912164;
      W_o[9,0] := -0.96086562;
      W_o[9,1] := -0.21338545;
      W_o[9,2] := -0.36878639;
      W_o[9,3] := -0.15249500;
      W_o[9,4] := -0.11614878;
      W_o[9,5] := -0.63825399;
      W_o[9,6] := -0.08493032;
      W_o[9,7] := -0.50577748;
      W_o[9,8] := -0.48369005;
      W_o[9,9] := 0.16791926;
      W_o[9,10] := -0.67517591;
      W_o[9,11] := -0.06844912;
      W_o[9,12] := -0.02455475;
      W_o[9,13] := 0.18983105;
      W_o[9,14] := 0.03197848;
      W_o[9,15] := -0.10859177;
      W_o[9,16] := -0.06121474;
      W_o[9,17] := 0.10381098;
      W_o[9,18] := -0.04804117;
      W_o[9,19] := -0.07395907;
      W_o[9,20] := -0.56294078;
      W_o[9,21] := 0.49253866;
      W_o[9,22] := -0.08418791;
      W_o[9,23] := 0.03632645;
      W_o[9,24] := -0.01930049;
      W_o[9,25] := 0.00721559;
      W_o[9,26] := 0.31399104;
      W_o[9,27] := 0.00363290;
      W_o[9,28] := 0.35762274;
      W_o[9,29] := 0.14383170;
      W_o[9,30] := 0.13138628;
      W_o[9,31] := -0.06635129;
      W_o[9,32] := 0.08883779;
      W_o[9,33] := 0.32405719;
      W_o[9,34] := -0.03502057;
      W_o[9,35] := -0.22428398;
      W_o[9,36] := -0.06680252;
      W_o[9,37] := -0.19686948;
      W_o[9,38] := 0.03372858;
      W_o[9,39] := -0.05063241;
      W_o[10,0] := -0.44047767;
      W_o[10,1] := -0.41061428;
      W_o[10,2] := 0.06679356;
      W_o[10,3] := 0.08232490;
      W_o[10,4] := 0.68651128;
      W_o[10,5] := 0.13447589;
      W_o[10,6] := -0.15820514;
      W_o[10,7] := -0.32401419;
      W_o[10,8] := 0.01493045;
      W_o[10,9] := 0.07515030;
      W_o[10,10] := -0.22708826;
      W_o[10,11] := -0.48697668;
      W_o[10,12] := -0.44020960;
      W_o[10,13] := -0.15198840;
      W_o[10,14] := -0.45878527;
      W_o[10,15] := -0.21131401;
      W_o[10,16] := -0.04725496;
      W_o[10,17] := -0.03169453;
      W_o[10,18] := 0.15397017;
      W_o[10,19] := -0.14169499;
      W_o[10,20] := 0.16080295;
      W_o[10,21] := -0.58566868;
      W_o[10,22] := -0.04027867;
      W_o[10,23] := -0.04846111;
      W_o[10,24] := 1.93909729;
      W_o[10,25] := 1.89536917;
      W_o[10,26] := -0.34381065;
      W_o[10,27] := -0.19164038;
      W_o[10,28] := 0.06696338;
      W_o[10,29] := 0.14391485;
      W_o[10,30] := -0.01906960;
      W_o[10,31] := 0.00395362;
      W_o[10,32] := 0.10876631;
      W_o[10,33] := 0.11656258;
      W_o[10,34] := 0.37426412;
      W_o[10,35] := 0.17253304;
      W_o[10,36] := 0.29803446;
      W_o[10,37] := 0.29228935;
      W_o[10,38] := 0.01999280;
      W_o[10,39] := 0.00505850;
      W_o[11,0] := 0.68408912;
      W_o[11,1] := 0.05380795;
      W_o[11,2] := 0.21208763;
      W_o[11,3] := -0.20944059;
      W_o[11,4] := 0.16949952;
      W_o[11,5] := -0.21931869;
      W_o[11,6] := -0.14467400;
      W_o[11,7] := -0.32249379;
      W_o[11,8] := 0.32598171;
      W_o[11,9] := -0.23611452;
      W_o[11,10] := -0.07394613;
      W_o[11,11] := -0.19434650;
      W_o[11,12] := 0.20823310;
      W_o[11,13] := -0.54425716;
      W_o[11,14] := -0.11235846;
      W_o[11,15] := -0.19877838;
      W_o[11,16] := 0.13296753;
      W_o[11,17] := 0.15389189;
      W_o[11,18] := 0.00750227;
      W_o[11,19] := 0.00651717;
      W_o[11,20] := -0.09164853;
      W_o[11,21] := 0.51982486;
      W_o[11,22] := 0.16873845;
      W_o[11,23] := -0.49257070;
      W_o[11,24] := -0.05849880;
      W_o[11,25] := 0.02633594;
      W_o[11,26] := 0.09369545;
      W_o[11,27] := -0.21366456;
      W_o[11,28] := 0.11514652;
      W_o[11,29] := 0.04365913;
      W_o[11,30] := 0.22134106;
      W_o[11,31] := 0.16536477;
      W_o[11,32] := -0.05712695;
      W_o[11,33] := 0.08705105;
      W_o[11,34] := 0.16276099;
      W_o[11,35] := -0.42817768;
      W_o[11,36] := 0.12246832;
      W_o[11,37] := -0.20113617;
      W_o[11,38] := 0.11593370;
      W_o[11,39] := -0.05348879;
      W_o[12,0] := -0.16644916;
      W_o[12,1] := -0.22179691;
      W_o[12,2] := -0.06963356;
      W_o[12,3] := 0.02390928;
      W_o[12,4] := -0.15694667;
      W_o[12,5] := 0.11342685;
      W_o[12,6] := 0.33777362;
      W_o[12,7] := -0.30824521;
      W_o[12,8] := -0.05667626;
      W_o[12,9] := -0.01847163;
      W_o[12,10] := 0.11112103;
      W_o[12,11] := -0.17032395;
      W_o[12,12] := -0.16411471;
      W_o[12,13] := -0.07482609;
      W_o[12,14] := -0.21282305;
      W_o[12,15] := -0.06134620;
      W_o[12,16] := 0.01745129;
      W_o[12,17] := -0.01394640;
      W_o[12,18] := 1.50527060;
      W_o[12,19] := -0.05658546;
      W_o[12,20] := -0.11261786;
      W_o[12,21] := -0.09813778;
      W_o[12,22] := 0.08243477;
      W_o[12,23] := 0.40823850;
      W_o[12,24] := -0.30796295;
      W_o[12,25] := -0.14412099;
      W_o[12,26] := 0.19181179;
      W_o[12,27] := 0.10502378;
      W_o[12,28] := 0.13072364;
      W_o[12,29] := 0.12108464;
      W_o[12,30] := 0.10646451;
      W_o[12,31] := -0.09400105;
      W_o[12,32] := -0.29639363;
      W_o[12,33] := 0.22136512;
      W_o[12,34] := -0.03096719;
      W_o[12,35] := 0.02072529;
      W_o[12,36] := -0.02478247;
      W_o[12,37] := -0.12082267;
      W_o[12,38] := -0.00598263;
      W_o[12,39] := -0.01071553;
      W_o[13,0] := -0.04834557;
      W_o[13,1] := 0.06634241;
      W_o[13,2] := -0.24370791;
      W_o[13,3] := 0.08637379;
      W_o[13,4] := -0.39779285;
      W_o[13,5] := 0.02139500;
      W_o[13,6] := 0.11640675;
      W_o[13,7] := 0.11385338;
      W_o[13,8] := -0.05518778;
      W_o[13,9] := 0.09104563;
      W_o[13,10] := 0.02279667;
      W_o[13,11] := -0.16343744;
      W_o[13,12] := -0.45273802;
      W_o[13,13] := -0.08252211;
      W_o[13,14] := -0.08964723;
      W_o[13,15] := -0.07374343;
      W_o[13,16] := -0.25515872;
      W_o[13,17] := -0.07434743;
      W_o[13,18] := 0.59073418;
      W_o[13,19] := 0.27197802;
      W_o[13,20] := -0.01829937;
      W_o[13,21] := 0.07717998;
      W_o[13,22] := 0.45007744;
      W_o[13,23] := 0.03504415;
      W_o[13,24] := 1.87039685;
      W_o[13,25] := 1.73898399;
      W_o[13,26] := 0.06699187;
      W_o[13,27] := -0.36609533;
      W_o[13,28] := 0.05306847;
      W_o[13,29] := 0.11336362;
      W_o[13,30] := 0.20086643;
      W_o[13,31] := -0.21461236;
      W_o[13,32] := -0.11377242;
      W_o[13,33] := -0.12958401;
      W_o[13,34] := 0.00505660;
      W_o[13,35] := -0.07748499;
      W_o[13,36] := -0.04069648;
      W_o[13,37] := 0.33590761;
      W_o[13,38] := 0.14594421;
      W_o[13,39] := -0.10981569;
      W_o[14,0] := -0.30323613;
      W_o[14,1] := -0.31149304;
      W_o[14,2] := 0.28586856;
      W_o[14,3] := 0.18452726;
      W_o[14,4] := 0.20233274;
      W_o[14,5] := -0.09256274;
      W_o[14,6] := -0.03783927;
      W_o[14,7] := 0.12692885;
      W_o[14,8] := -0.17600757;
      W_o[14,9] := 0.07501116;
      W_o[14,10] := -0.13759384;
      W_o[14,11] := 0.09564887;
      W_o[14,12] := 0.00343309;
      W_o[14,13] := 0.04607984;
      W_o[14,14] := -0.16881490;
      W_o[14,15] := -0.07940599;
      W_o[14,16] := -0.10241391;
      W_o[14,17] := -0.05080719;
      W_o[14,18] := 1.44254422;
      W_o[14,19] := -0.21181418;
      W_o[14,20] := 0.05755451;
      W_o[14,21] := 0.43047494;
      W_o[14,22] := -0.14185658;
      W_o[14,23] := 0.51635683;
      W_o[14,24] := 0.00273691;
      W_o[14,25] := 0.09392065;
      W_o[14,26] := -0.08311564;
      W_o[14,27] := 0.01820859;
      W_o[14,28] := 0.19468988;
      W_o[14,29] := 0.04482578;
      W_o[14,30] := -0.19548237;
      W_o[14,31] := -0.04979458;
      W_o[14,32] := 0.01701029;
      W_o[14,33] := 0.35701326;
      W_o[14,34] := 0.42355555;
      W_o[14,35] := -0.19557953;
      W_o[14,36] := 0.04753039;
      W_o[14,37] := 0.08129952;
      W_o[14,38] := -0.10219757;
      W_o[14,39] := 0.21446165;
      W_o[15,0] := -0.28090227;
      W_o[15,1] := 0.24640165;
      W_o[15,2] := -0.04431478;
      W_o[15,3] := 0.03227761;
      W_o[15,4] := -0.28705335;
      W_o[15,5] := 0.61719358;
      W_o[15,6] := -0.19619106;
      W_o[15,7] := -0.22106317;
      W_o[15,8] := -0.11724335;
      W_o[15,9] := 0.25582609;
      W_o[15,10] := -0.04176705;
      W_o[15,11] := 0.31498680;
      W_o[15,12] := 0.05772198;
      W_o[15,13] := 0.20806089;
      W_o[15,14] := -0.02345973;
      W_o[15,15] := 0.06730875;
      W_o[15,16] := 0.03451876;
      W_o[15,17] := -0.19311638;
      W_o[15,18] := -0.00410598;
      W_o[15,19] := -0.18493623;
      W_o[15,20] := -0.41258767;
      W_o[15,21] := -0.04694683;
      W_o[15,22] := -0.18209547;
      W_o[15,23] := -0.01441464;
      W_o[15,24] := -0.11699507;
      W_o[15,25] := -0.10582450;
      W_o[15,26] := 0.07790904;
      W_o[15,27] := -0.06042257;
      W_o[15,28] := 0.04504413;
      W_o[15,29] := 0.14734627;
      W_o[15,30] := -0.05427494;
      W_o[15,31] := 0.03112987;
      W_o[15,32] := 0.06163219;
      W_o[15,33] := 0.22637683;
      W_o[15,34] := 0.07694555;
      W_o[15,35] := -0.25882408;
      W_o[15,36] := 0.21838240;
      W_o[15,37] := -0.05452295;
      W_o[15,38] := 0.05332672;
      W_o[15,39] := 0.46538898;
      R_i[0,0] := -0.36683702;
      R_i[0,1] := -0.44737720;
      R_i[0,2] := 1.24589324;
      R_i[0,3] := 0.69412869;
      R_i[0,4] := 0.35085088;
      R_i[0,5] := -0.36259887;
      R_i[0,6] := 0.23951587;
      R_i[0,7] := 0.41614929;
      R_i[0,8] := 1.02476168;
      R_i[0,9] := 0.97401565;
      R_i[0,10] := 1.09034896;
      R_i[0,11] := -1.02841198;
      R_i[0,12] := -0.08663292;
      R_i[0,13] := 0.26691410;
      R_i[0,14] := -0.59099883;
      R_i[0,15] := 0.88828760;
      R_i[1,0] := -0.15458050;
      R_i[1,1] := 1.91954315;
      R_i[1,2] := -0.19880506;
      R_i[1,3] := -0.05338503;
      R_i[1,4] := 0.30228990;
      R_i[1,5] := -0.30340958;
      R_i[1,6] := 0.29198712;
      R_i[1,7] := -0.21350624;
      R_i[1,8] := -0.09833705;
      R_i[1,9] := 0.31499010;
      R_i[1,10] := -0.02912042;
      R_i[1,11] := 0.00149245;
      R_i[1,12] := 0.19466937;
      R_i[1,13] := 0.21224888;
      R_i[1,14] := -0.32503736;
      R_i[1,15] := -0.31977400;
      R_i[2,0] := -0.71105921;
      R_i[2,1] := -0.22115339;
      R_i[2,2] := -1.74462533;
      R_i[2,3] := -0.19147462;
      R_i[2,4] := 0.02834485;
      R_i[2,5] := 0.66907525;
      R_i[2,6] := 0.04054540;
      R_i[2,7] := -0.02422635;
      R_i[2,8] := 0.04692918;
      R_i[2,9] := 0.15513662;
      R_i[2,10] := -0.05168056;
      R_i[2,11] := -0.07468271;
      R_i[2,12] := -0.57621449;
      R_i[2,13] := -0.14785919;
      R_i[2,14] := 0.40508196;
      R_i[2,15] := 0.20491433;
      R_i[3,0] := 0.30087462;
      R_i[3,1] := 0.81402808;
      R_i[3,2] := -0.53180295;
      R_i[3,3] := -2.29824114;
      R_i[3,4] := 0.49502930;
      R_i[3,5] := 0.07546997;
      R_i[3,6] := -0.41725859;
      R_i[3,7] := 0.29847994;
      R_i[3,8] := 0.09713065;
      R_i[3,9] := -0.08287358;
      R_i[3,10] := 0.16965586;
      R_i[3,11] := -0.26217785;
      R_i[3,12] := 0.14900748;
      R_i[3,13] := 0.36093932;
      R_i[3,14] := -0.33660060;
      R_i[3,15] := -0.90025556;
      R_i[4,0] := -3.00713706;
      R_i[4,1] := -0.16220070;
      R_i[4,2] := 0.86550975;
      R_i[4,3] := 0.14306493;
      R_i[4,4] := -1.69561899;
      R_i[4,5] := -0.23536262;
      R_i[4,6] := 1.44078171;
      R_i[4,7] := 0.40745640;
      R_i[4,8] := 0.84672201;
      R_i[4,9] := 0.61333311;
      R_i[4,10] := -0.13707401;
      R_i[4,11] := -0.82632464;
      R_i[4,12] := 0.75525576;
      R_i[4,13] := 0.10271102;
      R_i[4,14] := -0.39098045;
      R_i[4,15] := -0.34274298;
      R_i[5,0] := 0.29963374;
      R_i[5,1] := 0.10178780;
      R_i[5,2] := 0.32936281;
      R_i[5,3] := 0.29712185;
      R_i[5,4] := 0.21390122;
      R_i[5,5] := -0.24001811;
      R_i[5,6] := 0.04780090;
      R_i[5,7] := -0.06073575;
      R_i[5,8] := -0.07838094;
      R_i[5,9] := -0.04620231;
      R_i[5,10] := 0.43323347;
      R_i[5,11] := -0.42312637;
      R_i[5,12] := -0.02658233;
      R_i[5,13] := -0.26356259;
      R_i[5,14] := 0.06192940;
      R_i[5,15] := -0.13695642;
      R_i[6,0] := -0.67857140;
      R_i[6,1] := -0.50468159;
      R_i[6,2] := 0.26149645;
      R_i[6,3] := -0.23731886;
      R_i[6,4] := 0.32474071;
      R_i[6,5] := -1.04019964;
      R_i[6,6] := -0.14901595;
      R_i[6,7] := 0.48365265;
      R_i[6,8] := -0.06066033;
      R_i[6,9] := -0.61287755;
      R_i[6,10] := -0.44098693;
      R_i[6,11] := 0.17185783;
      R_i[6,12] := -0.02349554;
      R_i[6,13] := -0.49048305;
      R_i[6,14] := 0.24112639;
      R_i[6,15] := -0.11388259;
      R_i[7,0] := 0.19145711;
      R_i[7,1] := -0.52626193;
      R_i[7,2] := 0.14510420;
      R_i[7,3] := -0.35204259;
      R_i[7,4] := 0.86173880;
      R_i[7,5] := 0.70634562;
      R_i[7,6] := 0.08693185;
      R_i[7,7] := -1.86060202;
      R_i[7,8] := -0.48649496;
      R_i[7,9] := 0.36919993;
      R_i[7,10] := 0.12250333;
      R_i[7,11] := 0.22951156;
      R_i[7,12] := 0.02786869;
      R_i[7,13] := 0.52622157;
      R_i[7,14] := 0.56637853;
      R_i[7,15] := -0.16136852;
      R_i[8,0] := -0.53185570;
      R_i[8,1] := -0.04072466;
      R_i[8,2] := -0.14449374;
      R_i[8,3] := -0.13692714;
      R_i[8,4] := 0.82504284;
      R_i[8,5] := 0.19167326;
      R_i[8,6] := 1.67909050;
      R_i[8,7] := 0.29732254;
      R_i[8,8] := -1.54010010;
      R_i[8,9] := 0.05109580;
      R_i[8,10] := 0.31016925;
      R_i[8,11] := -0.34457940;
      R_i[8,12] := -0.33437556;
      R_i[8,13] := 0.09498347;
      R_i[8,14] := -0.53118694;
      R_i[8,15] := -0.08159891;
      R_i[9,0] := -0.15789132;
      R_i[9,1] := 0.21440165;
      R_i[9,2] := -0.11797124;
      R_i[9,3] := -0.31671742;
      R_i[9,4] := 0.13391078;
      R_i[9,5] := -0.04241018;
      R_i[9,6] := 0.13570282;
      R_i[9,7] := -0.37446287;
      R_i[9,8] := 0.06697363;
      R_i[9,9] := -0.31501204;
      R_i[9,10] := 0.08753272;
      R_i[9,11] := 0.14745103;
      R_i[9,12] := 0.25471240;
      R_i[9,13] := -0.00752171;
      R_i[9,14] := -0.13687773;
      R_i[9,15] := -0.20334294;
      R_i[10,0] := 0.10601140;
      R_i[10,1] := 0.33716449;
      R_i[10,2] := -0.28345254;
      R_i[10,3] := -0.08123855;
      R_i[10,4] := 0.65765005;
      R_i[10,5] := -0.16018872;
      R_i[10,6] := 0.66867888;
      R_i[10,7] := 0.05066697;
      R_i[10,8] := -0.26125985;
      R_i[10,9] := 0.06136491;
      R_i[10,10] := -0.07193215;
      R_i[10,11] := -0.00455745;
      R_i[10,12] := 0.50109005;
      R_i[10,13] := -0.34902012;
      R_i[10,14] := -0.10270999;
      R_i[10,15] := -0.27994797;
      R_i[11,0] := 0.16313595;
      R_i[11,1] := -0.19938010;
      R_i[11,2] := 0.06057022;
      R_i[11,3] := -0.01475503;
      R_i[11,4] := 0.54161280;
      R_i[11,5] := -0.03717137;
      R_i[11,6] := 0.43041891;
      R_i[11,7] := 0.10488611;
      R_i[11,8] := -0.33726332;
      R_i[11,9] := -0.35081905;
      R_i[11,10] := -0.12337096;
      R_i[11,11] := 0.50985360;
      R_i[11,12] := 0.00059109;
      R_i[11,13] := 0.11848055;
      R_i[11,14] := -0.06023524;
      R_i[11,15] := 0.00647274;
      R_i[12,0] := -1.13358891;
      R_i[12,1] := 0.25045577;
      R_i[12,2] := -0.72799140;
      R_i[12,3] := -0.28028357;
      R_i[12,4] := -0.25076982;
      R_i[12,5] := 0.41504830;
      R_i[12,6] := 0.96340883;
      R_i[12,7] := 0.06510375;
      R_i[12,8] := 0.33402908;
      R_i[12,9] := 0.07096598;
      R_i[12,10] := 0.59124023;
      R_i[12,11] := -0.12774691;
      R_i[12,12] := 2.18120933;
      R_i[12,13] := -0.54086334;
      R_i[12,14] := 0.75623906;
      R_i[12,15] := -0.67408884;
      R_i[13,0] := -0.85261506;
      R_i[13,1] := 0.17393038;
      R_i[13,2] := -0.10425876;
      R_i[13,3] := -0.27151591;
      R_i[13,4] := -0.57615143;
      R_i[13,5] := 0.06762128;
      R_i[13,6] := 0.17267182;
      R_i[13,7] := 0.58947426;
      R_i[13,8] := -0.37534830;
      R_i[13,9] := -0.18215351;
      R_i[13,10] := -0.33110857;
      R_i[13,11] := -0.27655941;
      R_i[13,12] := -0.40030205;
      R_i[13,13] := 1.32292378;
      R_i[13,14] := 0.21090908;
      R_i[13,15] := -0.05352690;
      R_i[14,0] := 0.03172403;
      R_i[14,1] := -0.48991668;
      R_i[14,2] := -0.05704284;
      R_i[14,3] := 0.11988008;
      R_i[14,4] := 0.17805719;
      R_i[14,5] := 0.23852935;
      R_i[14,6] := 0.12931433;
      R_i[14,7] := -0.03777663;
      R_i[14,8] := 0.07517263;
      R_i[14,9] := -0.03596207;
      R_i[14,10] := 0.04425231;
      R_i[14,11] := -0.36268836;
      R_i[14,12] := -0.02361461;
      R_i[14,13] := 0.16448504;
      R_i[14,14] := -0.30058336;
      R_i[14,15] := -0.16361728;
      R_i[15,0] := 0.74356866;
      R_i[15,1] := 0.25941604;
      R_i[15,2] := -0.17731465;
      R_i[15,3] := -0.18815078;
      R_i[15,4] := 0.48738170;
      R_i[15,5] := 0.13013434;
      R_i[15,6] := -0.12726560;
      R_i[15,7] := 0.27749133;
      R_i[15,8] := 0.35979366;
      R_i[15,9] := 0.25837585;
      R_i[15,10] := -0.69103974;
      R_i[15,11] := -0.36489427;
      R_i[15,12] := 0.03232842;
      R_i[15,13] := 0.32356966;
      R_i[15,14] := -0.20295747;
      R_i[15,15] := -0.26835045;
      R_f[0,0] := 0.07153955;
      R_f[0,1] := -0.59087461;
      R_f[0,2] := 0.49619547;
      R_f[0,3] := 0.07594358;
      R_f[0,4] := 0.24425711;
      R_f[0,5] := 0.14149903;
      R_f[0,6] := -0.09984472;
      R_f[0,7] := 0.10858753;
      R_f[0,8] := 0.25852686;
      R_f[0,9] := 0.16836661;
      R_f[0,10] := -0.49937955;
      R_f[0,11] := 0.18961865;
      R_f[0,12] := -0.49092764;
      R_f[0,13] := 0.15820153;
      R_f[0,14] := -0.06552398;
      R_f[0,15] := -0.14661682;
      R_f[1,0] := -0.05355694;
      R_f[1,1] := 1.92975557;
      R_f[1,2] := 0.27318946;
      R_f[1,3] := 0.94045126;
      R_f[1,4] := 0.01676022;
      R_f[1,5] := 0.07051807;
      R_f[1,6] := 0.18478443;
      R_f[1,7] := -0.37505114;
      R_f[1,8] := 0.09433642;
      R_f[1,9] := 0.10628120;
      R_f[1,10] := -0.30447745;
      R_f[1,11] := 0.35159656;
      R_f[1,12] := 0.45133221;
      R_f[1,13] := -0.04233953;
      R_f[1,14] := 0.77227736;
      R_f[1,15] := 0.55623603;
      R_f[2,0] := -0.29655850;
      R_f[2,1] := 0.87102282;
      R_f[2,2] := -1.04400361;
      R_f[2,3] := -0.26446375;
      R_f[2,4] := 0.30872551;
      R_f[2,5] := 0.53280818;
      R_f[2,6] := 0.08578387;
      R_f[2,7] := 0.27742198;
      R_f[2,8] := 0.32091269;
      R_f[2,9] := -0.35130039;
      R_f[2,10] := 0.13140900;
      R_f[2,11] := -0.01945328;
      R_f[2,12] := 0.62961471;
      R_f[2,13] := -0.47139388;
      R_f[2,14] := 0.81306297;
      R_f[2,15] := 0.06325053;
      R_f[3,0] := -0.52896017;
      R_f[3,1] := 0.37202662;
      R_f[3,2] := -0.03908378;
      R_f[3,3] := -1.92155027;
      R_f[3,4] := -0.15915719;
      R_f[3,5] := 0.04583488;
      R_f[3,6] := 0.26791275;
      R_f[3,7] := 0.17511773;
      R_f[3,8] := -0.40435636;
      R_f[3,9] := -0.03977980;
      R_f[3,10] := 0.47443610;
      R_f[3,11] := -0.07829616;
      R_f[3,12] := 0.21981125;
      R_f[3,13] := 0.11550741;
      R_f[3,14] := 0.28196028;
      R_f[3,15] := -0.41792643;
      R_f[4,0] := -0.16650143;
      R_f[4,1] := -0.89877087;
      R_f[4,2] := 0.86069864;
      R_f[4,3] := 0.30464059;
      R_f[4,4] := -0.05939668;
      R_f[4,5] := 0.25487947;
      R_f[4,6] := 1.13254857;
      R_f[4,7] := -0.40170091;
      R_f[4,8] := -0.60228431;
      R_f[4,9] := 0.17544644;
      R_f[4,10] := -0.03666126;
      R_f[4,11] := -1.09364593;
      R_f[4,12] := 0.14268741;
      R_f[4,13] := -0.03543003;
      R_f[4,14] := 0.25145757;
      R_f[4,15] := 0.06923623;
      R_f[5,0] := 0.07152445;
      R_f[5,1] := -0.93268287;
      R_f[5,2] := 0.96183014;
      R_f[5,3] := 0.34152153;
      R_f[5,4] := 0.11259452;
      R_f[5,5] := 0.13736168;
      R_f[5,6] := 0.45562023;
      R_f[5,7] := -0.12320174;
      R_f[5,8] := -0.39810219;
      R_f[5,9] := -0.61624128;
      R_f[5,10] := -0.15761711;
      R_f[5,11] := -0.32445639;
      R_f[5,12] := -0.21541518;
      R_f[5,13] := -0.01548673;
      R_f[5,14] := -0.18224493;
      R_f[5,15] := 0.16112094;
      R_f[6,0] := -0.01400591;
      R_f[6,1] := -1.15473711;
      R_f[6,2] := 0.46569550;
      R_f[6,3] := 0.35570300;
      R_f[6,4] := 0.64884621;
      R_f[6,5] := 0.68359298;
      R_f[6,6] := -0.61912656;
      R_f[6,7] := -0.18728444;
      R_f[6,8] := -1.13906693;
      R_f[6,9] := -0.60935068;
      R_f[6,10] := -0.23855972;
      R_f[6,11] := -0.49719852;
      R_f[6,12] := 0.25523233;
      R_f[6,13] := -1.26516819;
      R_f[6,14] := -0.21763113;
      R_f[6,15] := 0.12647545;
      R_f[7,0] := 2.03078747;
      R_f[7,1] := -0.76834255;
      R_f[7,2] := 0.61253548;
      R_f[7,3] := 0.39429587;
      R_f[7,4] := -0.30242923;
      R_f[7,5] := 2.34057760;
      R_f[7,6] := 2.17685127;
      R_f[7,7] := -2.06056809;
      R_f[7,8] := -1.78221929;
      R_f[7,9] := 0.36663124;
      R_f[7,10] := 0.72593582;
      R_f[7,11] := -0.06118135;
      R_f[7,12] := -1.00646436;
      R_f[7,13] := 1.82777369;
      R_f[7,14] := 0.38762328;
      R_f[7,15] := 0.51006883;
      R_f[8,0] := -0.06902416;
      R_f[8,1] := -1.26130819;
      R_f[8,2] := 0.95632678;
      R_f[8,3] := -0.08877252;
      R_f[8,4] := 0.02389756;
      R_f[8,5] := -0.23528144;
      R_f[8,6] := 0.16436763;
      R_f[8,7] := -0.05826518;
      R_f[8,8] := -2.04791641;
      R_f[8,9] := -0.42510942;
      R_f[8,10] := -0.24232592;
      R_f[8,11] := -0.51980168;
      R_f[8,12] := -0.14773984;
      R_f[8,13] := -0.49321669;
      R_f[8,14] := 0.28463793;
      R_f[8,15] := -0.21783537;
      R_f[9,0] := -0.13374837;
      R_f[9,1] := -1.17639554;
      R_f[9,2] := 0.12627633;
      R_f[9,3] := 0.06300414;
      R_f[9,4] := 0.01875936;
      R_f[9,5] := -0.21104464;
      R_f[9,6] := -0.02009901;
      R_f[9,7] := -0.71492696;
      R_f[9,8] := -0.88293582;
      R_f[9,9] := -1.22890174;
      R_f[9,10] := -0.09347305;
      R_f[9,11] := -0.60869575;
      R_f[9,12] := -0.13751322;
      R_f[9,13] := 0.35621238;
      R_f[9,14] := 0.79695553;
      R_f[9,15] := 1.19073606;
      R_f[10,0] := -0.29936871;
      R_f[10,1] := -0.73769796;
      R_f[10,2] := 0.06686691;
      R_f[10,3] := 0.29226211;
      R_f[10,4] := -0.24629065;
      R_f[10,5] := 0.97109705;
      R_f[10,6] := 0.28993571;
      R_f[10,7] := -0.64702898;
      R_f[10,8] := -0.33609614;
      R_f[10,9] := 0.15665323;
      R_f[10,10] := 0.20275173;
      R_f[10,11] := 0.28188258;
      R_f[10,12] := -0.35766971;
      R_f[10,13] := -0.45825234;
      R_f[10,14] := 0.59465575;
      R_f[10,15] := -0.09009458;
      R_f[11,0] := -0.06559964;
      R_f[11,1] := -0.34416181;
      R_f[11,2] := 0.06520309;
      R_f[11,3] := -0.01709294;
      R_f[11,4] := -0.44365394;
      R_f[11,5] := 0.10967853;
      R_f[11,6] := 0.18147334;
      R_f[11,7] := -0.28511751;
      R_f[11,8] := 0.30923906;
      R_f[11,9] := 0.29513508;
      R_f[11,10] := -0.18808335;
      R_f[11,11] := -0.27482635;
      R_f[11,12] := 0.11784156;
      R_f[11,13] := 0.21471596;
      R_f[11,14] := 0.22612707;
      R_f[11,15] := 0.32492065;
      R_f[12,0] := 0.66689140;
      R_f[12,1] := -0.79796457;
      R_f[12,2] := 0.76750970;
      R_f[12,3] := 0.37235740;
      R_f[12,4] := -0.73377728;
      R_f[12,5] := -0.09779347;
      R_f[12,6] := 0.12647966;
      R_f[12,7] := -0.62336546;
      R_f[12,8] := 0.00648065;
      R_f[12,9] := -0.26842323;
      R_f[12,10] := 1.69255817;
      R_f[12,11] := 0.01504949;
      R_f[12,12] := 0.38201123;
      R_f[12,13] := -0.21126585;
      R_f[12,14] := 0.79340529;
      R_f[12,15] := -0.67332441;
      R_f[13,0] := 0.18675253;
      R_f[13,1] := 0.29937005;
      R_f[13,2] := 0.15947086;
      R_f[13,3] := 0.30692375;
      R_f[13,4] := -0.11816163;
      R_f[13,5] := 0.34528661;
      R_f[13,6] := -0.42399773;
      R_f[13,7] := -0.11187272;
      R_f[13,8] := -0.08543108;
      R_f[13,9] := 0.45360404;
      R_f[13,10] := 0.08977752;
      R_f[13,11] := -0.08927725;
      R_f[13,12] := 0.74914813;
      R_f[13,13] := 0.32484278;
      R_f[13,14] := 0.27966246;
      R_f[13,15] := 0.64148533;
      R_f[14,0] := 0.00067597;
      R_f[14,1] := 0.03178573;
      R_f[14,2] := 0.24933998;
      R_f[14,3] := -0.18668689;
      R_f[14,4] := 0.22304797;
      R_f[14,5] := -0.05844809;
      R_f[14,6] := 0.01542039;
      R_f[14,7] := -0.07623729;
      R_f[14,8] := -0.19314471;
      R_f[14,9] := -0.21212263;
      R_f[14,10] := 0.23236075;
      R_f[14,11] := -0.57485098;
      R_f[14,12] := 0.46047559;
      R_f[14,13] := -0.00148298;
      R_f[14,14] := -0.21503349;
      R_f[14,15] := -0.12761565;
      R_f[15,0] := 0.23568556;
      R_f[15,1] := -0.97643197;
      R_f[15,2] := 0.21373613;
      R_f[15,3] := 0.39719129;
      R_f[15,4] := -0.24737620;
      R_f[15,5] := 0.22643280;
      R_f[15,6] := 0.64512557;
      R_f[15,7] := 0.19389327;
      R_f[15,8] := -0.60527653;
      R_f[15,9] := -0.22903773;
      R_f[15,10] := -0.28841779;
      R_f[15,11] := -0.52285588;
      R_f[15,12] := -0.59739178;
      R_f[15,13] := -0.20141296;
      R_f[15,14] := 0.29787028;
      R_f[15,15] := -1.29604101;
      R_g[0,0] := -1.70048869;
      R_g[0,1] := -0.02498771;
      R_g[0,2] := 0.05516972;
      R_g[0,3] := 0.22662289;
      R_g[0,4] := -0.23178743;
      R_g[0,5] := 0.13714461;
      R_g[0,6] := 0.16423392;
      R_g[0,7] := -0.08702778;
      R_g[0,8] := -0.05017116;
      R_g[0,9] := 0.03059242;
      R_g[0,10] := 0.00949551;
      R_g[0,11] := -0.08035634;
      R_g[0,12] := 0.07701789;
      R_g[0,13] := -0.13365406;
      R_g[0,14] := -0.11454831;
      R_g[0,15] := 0.32707965;
      R_g[1,0] := 0.00018709;
      R_g[1,1] := -1.38878047;
      R_g[1,2] := -0.24736334;
      R_g[1,3] := -0.08500341;
      R_g[1,4] := 0.03873841;
      R_g[1,5] := -0.00933929;
      R_g[1,6] := 0.01160030;
      R_g[1,7] := -0.06713413;
      R_g[1,8] := 0.03234413;
      R_g[1,9] := 0.27781528;
      R_g[1,10] := -0.22306302;
      R_g[1,11] := -0.29338247;
      R_g[1,12] := 0.30125844;
      R_g[1,13] := 0.38746142;
      R_g[1,14] := -0.23414122;
      R_g[1,15] := -0.22076719;
      R_g[2,0] := -0.15139687;
      R_g[2,1] := 0.14425665;
      R_g[2,2] := -0.51542902;
      R_g[2,3] := -0.12809730;
      R_g[2,4] := 0.04208002;
      R_g[2,5] := -0.07483902;
      R_g[2,6] := -0.00554008;
      R_g[2,7] := 0.23140340;
      R_g[2,8] := -0.06807555;
      R_g[2,9] := 0.01600222;
      R_g[2,10] := 0.06458747;
      R_g[2,11] := -0.45057061;
      R_g[2,12] := 0.26487321;
      R_g[2,13] := 0.28997588;
      R_g[2,14] := -0.39954144;
      R_g[2,15] := -0.56048697;
      R_g[3,0] := 0.22866221;
      R_g[3,1] := 0.67594492;
      R_g[3,2] := -0.40921754;
      R_g[3,3] := -1.74979711;
      R_g[3,4] := 0.11497030;
      R_g[3,5] := -0.06326534;
      R_g[3,6] := -0.10878199;
      R_g[3,7] := 0.01786116;
      R_g[3,8] := 0.05380635;
      R_g[3,9] := 0.03915313;
      R_g[3,10] := -0.08796055;
      R_g[3,11] := -0.60486305;
      R_g[3,12] := 0.14022473;
      R_g[3,13] := 0.09025718;
      R_g[3,14] := -0.17233410;
      R_g[3,15] := -0.83184385;
      R_g[4,0] := 0.11942312;
      R_g[4,1] := -0.03900880;
      R_g[4,2] := 0.22554153;
      R_g[4,3] := 0.24997710;
      R_g[4,4] := -2.11677217;
      R_g[4,5] := 0.18121429;
      R_g[4,6] := 0.03432639;
      R_g[4,7] := -0.15975657;
      R_g[4,8] := -0.03747511;
      R_g[4,9] := 0.06238879;
      R_g[4,10] := -0.13933714;
      R_g[4,11] := -0.26897860;
      R_g[4,12] := -0.11694002;
